(* IEC 61131-3 sources: daoli-st-library/DL_Device (part 32) *)

(* ---- FB_DL_StarDeltaMotor.st ---- *)
(*==============================================================================
 * 组件名称 (Component)  : FB_DL_StarDeltaMotor
 * 所属子库 (Sublibrary) : DL_Device
 * 当前版本 (Version)    : 1.0.1
 * 兼容性   (Platform)   : CODESYS 3.5 / TwinCAT 3 / 汇川 InoProShop / Machine Expert
 *                         仅依赖 Standard.library（TON / R_TRIG），零厂商方言
 * 分类     (Category)   : 设备执行器功能块（Function Block，无接口实现）
 * 功能简述 (Function)   : 星三角降压启动电机控制（三接触器）。星形降压启动
 *                         （起动力矩约三分之一）→ 星角切换死区互锁（星线圈
 *                         分断后方允许角线圈吸合）→ 三角形全压运行；三路
 *                         接触器指令-反馈校验窗（拒动保护）、运行失反馈
 *                         脱扣、热继过载锁存、重启抑制冷却（沿用
 *                         FB_DL_DolMotor 参数范式）；星角输出互斥出口
 *                         断言 + 反馈互锁冲突监视；状态机复用既有
 *                         E_DL_MotorState（禁止重定义），ENUM + CASE + ELSE
 *                         兜底。
 * 开源溯源 (Origin)     : 来源标签 lbp-basic-process / lbp-device
 *                         （RAW_NOTES_R6 S-1 + S-5：星三角降压启动时序、
 *                         星角切换死区时间互锁、三接触器反馈校验等行业
 *                         公知工程惯例，公开教学资料，仅借鉴通用工程语义；
 *                         状态机、死区互锁实现、故障码按本库红线独立设计，
 *                         clean-room 未复制源码）。
 * 红线自检 (Redline)    : R1 零全局变量表/外部变量引用 ✓｜R2 零物理 IO 地址 ✓
 *                         R3 纯 IEC 61131-3 ✓｜R4 防越界/互斥断言 ✓
 *                         R5 全变量中英双语同行注释 ✓｜R6 ENUM+CASE+ELSE ✓
 *                         R7 七个定时器/边缘实例主体最前部无条件刷新 ✓
 * 公约遵循 (Convention) : 0.1/R23 本块为纯事件型状态机（BOOL 指令/反馈 +
 *                         TIME 参数，无积分/滤波类连续量同步语义），免首扫，
 *                         无内部初始化标志。
 *                         0.7 故障码段位 16#0003_xxxx：【故障级】0003_0240
 *                         主接触器拒动 / 0003_0241 星接触器拒动 / 0003_0242
 *                         星接触器分断失败（角拒动码位承接，见偏离③）/
 *                         0003_0243 星角互斥冲突 / 0003_0244 运行失反馈
 *                         脱扣 / 0003_0245 过载锁存 / 0003_0246 星角转换
 *                         失败（角接触器窗内未吸合），全部 R15 锁存仅复位
 *                         可清；【信息级】0003_0208 重启抑制期启动拒绝
 *                         （沿用 FB_DL_DolMotor 既有同义码位，终审裁定统
 *                         一双电机族口径；仅写 uErrorId，不进 bFault，0.2
 *                         公约）。
 * 偏离留档 (Deviation)  : 依 R11 头注释留档，共 3 条：
 *                         ① 信息级码：规格原分配 0003_0102，经与子库
 *                           VERSION.md 故障码表核对，R5 已占用 0102~0104
 *                           （AnalogTransmitter）；且重启抑制拒绝语义在
 *                           FB_DL_DolMotor 已有信息级码位 0003_0208——
 *                           终审裁定同库同语义不设双码，本块改用 0208
 *                           （0105 空置不分配），与规格原意"沿用 DolMotor
 *                           口径"完全一致。
 *                         ② 规格中 0003_0242（角接触器拒动）与 0003_0246
 *                           （星角转换失败）对"死区满后角接触器窗内未吸合"
 *                           同事件重叠；本实现将 0246 用于规格明示的角接触
 *                           器窗内未吸合，0242 承接转换窗口内星接触器反馈
 *                           未按时分断（星粘连/拒分）的互锁异常，两码位
 *                           各自可测。
 *                         ③ 重启抑制冷却计时采用 TON（本库 Standard.library
 *                           既有范式，DolMotor 同口径），无 CPU 钟依赖。
 * 修订历史 (Revision)   :
 *   2026-11-15  v1.0.0  首版入库（R6 轮 · DL_Device 阀门/驱动族深化）
 *   2026-11-15  v1.0.1  终审修复【逻辑级】重启抑制信息级码双码归一：原分配
 *                       0003_0105 与 FB_DL_DolMotor 既有同义码 0003_0208
 *                       重复（同库同语义双码会致 HMI 报警分组重复映射），
 *                       改用 0208 统一口径。引脚契约零变更。
 *============================================================================*)
FUNCTION_BLOCK FB_DL_StarDeltaMotor
VAR_INPUT
    bCmdStart        : BOOL;            // 启动指令（Start command），上升沿生效 / Start command, rising edge effective
    bCmdStop         : BOOL;            // 停止指令（Stop command），电平生效 / Stop command, level effective
    bFbMain          : BOOL;            // 主接触器反馈（Main contactor feedback），TRUE=吸合 / Main contactor feedback, TRUE = picked up
    bFbStar          : BOOL;            // 星形接触器反馈（Star contactor feedback），TRUE=吸合 / Star contactor feedback, TRUE = picked up
    bFbDelta         : BOOL;            // 三角形接触器反馈（Delta contactor feedback），TRUE=吸合 / Delta contactor feedback, TRUE = picked up
    bThermalOverload : BOOL;            // 热继电器过载信号（Thermal overload trip），TRUE=过载 / Thermal overload trip, TRUE = overloaded
    bPermitStart     : BOOL;            // 启动允许联锁（Start permit），TRUE=允许 / Start permit interlock, TRUE = start allowed
    tStarTime        : TIME := T#5S;    // 星形运行时间（Star run time），按负载实测加速时间整定 / Star run time, tune per measured load acceleration
    tDeadTime        : TIME := T#100MS; // 星角转换死区时间（Transition dead time），域 50~200MS，星分断后角方可吸合 / Transition dead time 50..200 ms, star must drop before delta picks up
    tFbWindow        : TIME := T#500MS; // 指令-反馈校验窗口（Feedback check window），T#0S=免校验 / Feedback check window, T#0S disables the check
    tRestartInhibit  : TIME := T#60S;   // 重启抑制冷却时间（Restart inhibit），停机后冷却期内拒绝启动 / Restart inhibit cooling time after stop
    bReset           : BOOL;            // 故障复位（Fault reset），上升沿生效 / Fault reset, rising edge effective
END_VAR

VAR_OUTPUT
    bMainContactor   : BOOL;            // 主接触器线圈输出（Main contactor coil），星形与运行期全程吸合 / Main contactor coil, closed through star and run phases
    bStarContactor   : BOOL;            // 星形接触器线圈输出（Star contactor coil），仅星形降压段吸合 / Star contactor coil, closed only in star phase
    bDeltaContactor  : BOOL;            // 三角形接触器线圈输出（Delta contactor coil），死区满后吸合 / Delta contactor coil, closed after dead time
    eState           : E_DL_MotorState; // 当前状态机状态（Current state），复用既有枚举 / Current state, reuses existing enum
    bRunning         : BOOL;            // 运行反馈（Running feedback），角接触器吸合确认 / Running feedback, confirmed by delta contactor
    bFault           : BOOL;            // 故障锁存中（Fault latched），TRUE=需复位（含过载脱扣）/ Fault latched, TRUE requires reset (incl. overload trip)
    uErrorId         : UDINT;           // 末次故障码（Last error code），0=无故障，段位 16#0003_xxxx / Last error code, 0 = none, family 16#0003_xxxx
    bRestartInhibit  : BOOL;            // 重启抑制激活中（Restart inhibit active），TRUE=冷却期拒绝启动 / Restart inhibit active, TRUE = starts refused
    bStarPhase       : BOOL;            // 星形阶段指示（Star phase active），调试/HMI 用 / Star phase indicator for debug and HMI
    uStartCount      : UDINT;           // 累计启动次数（Start count），每次受理启动 +1 / Total start count, incremented per accepted start
END_VAR

VAR
    _eState           : E_DL_MotorState := E_DL_MotorState.eIdle; // 内部状态机步序（Internal state step）/ Internal state step
    _bFaultLatch      : BOOL;           // 故障锁存标志（Fault latch flag），仅复位清除 / Fault latch flag, cleared only by reset
    _uErrorIdInt      : UDINT;          // 内部故障码寄存（Internal error register），故障级与信息级共用 / Internal error register, fault and info codes share it
    _bDeadZone        : BOOL;           // 星角转换死区子相位（Star-delta dead-zone sub-phase），星形态内二段 / Dead-zone sub-phase inside starting state
    _bDeltaCmd        : BOOL;           // 角接触器指令已发出（Delta command issued），转换校验窗运行中 / Delta command issued, check window running
    _bCooling         : BOOL;           // 冷却计时进行中（Cooling timing active）/ Cooling timer run request flag
    _bRestartInhAct   : BOOL;           // 重启抑制激活内部寄存（Internal restart inhibit register）/ Internal restart inhibit register
    _bFbWinEn         : BOOL;           // 反馈校验窗使能（Feedback window enable），窗口参数大于零有效 / Feedback window enable, active when window above zero
    _bInFbWin         : BOOL;           // 主/星反馈窗计时条件（Main/star window timing condition）/ Timing condition of main and star window
    _bInStarTime      : BOOL;           // 星形运行计时条件（Star run timing condition）/ Timing condition of star run timer
    _bInDeadTime      : BOOL;           // 死区计时条件（Dead time timing condition）/ Timing condition of dead time timer
    _bInDeltaWin      : BOOL;           // 角反馈窗计时条件（Delta window timing condition）/ Timing condition of delta window
    _bInRunningSt     : BOOL;           // 运行态判定中间量（Running-state test intermediate） / Running-state test intermediate
    _fbTrigStart      : R_TRIG;         // 引脚启动指令上升沿（Pin start command edge）/ Pin start command rising edge
    _fbTrigReset      : R_TRIG;         // 引脚复位上升沿（Pin reset edge）/ Pin reset rising edge
    _fbTonFbWin       : TON;            // 主/星接触器反馈校验窗定时器（Main and star feedback window timer）/ Main and star feedback window timer
    _fbTonStarTime    : TON;            // 星形运行时间定时器（Star run time timer）/ Star run time timer
    _fbTonDeadTime    : TON;            // 星角转换死区定时器（Transition dead time timer）/ Transition dead time timer
    _fbTonDeltaWin    : TON;            // 角接触器反馈校验窗定时器（Delta feedback window timer）/ Delta feedback window timer
    _fbTonRestartInh  : TON;            // 重启抑制冷却定时器（Restart inhibit cooling timer）/ Restart inhibit cooling timer
END_VAR

// ============================================================================
// 段 1｜定时器与边缘检测实例无条件周期刷新（R7：严禁置于 IF/CASE 分支内）
//      Unconditional per-cycle refresh of all timer and edge instances (R7)
// ============================================================================
_fbTrigStart(CLK := bCmdStart);
_fbTrigReset(CLK := bReset);
_bFbWinEn := (tFbWindow > T#0S);      // 窗口为零 = 免校验（Zero window = check disabled）
_bInFbWin := (_eState = E_DL_MotorState.eStarting) AND (NOT _bDeadZone) AND _bFbWinEn; // 启动段主/星校验窗（Starting phase main and star window）
_bInStarTime := (_eState = E_DL_MotorState.eStarting) AND (NOT _bDeadZone); // 星形段计时（Star phase timing）
_bInDeadTime := (_eState = E_DL_MotorState.eStarting) AND _bDeadZone AND (NOT _bDeltaCmd); // 死区段计时（Dead-zone timing）
_bInDeltaWin := (_eState = E_DL_MotorState.eStarting) AND _bDeadZone AND _bDeltaCmd AND (NOT bFbDelta) AND _bFbWinEn; // 角校验窗（Delta check window）
_fbTonFbWin(IN := _bInFbWin, PT := tFbWindow);
_fbTonStarTime(IN := _bInStarTime, PT := tStarTime);
_fbTonDeadTime(IN := _bInDeadTime, PT := tDeadTime);
_fbTonDeltaWin(IN := _bInDeltaWin, PT := tFbWindow);
_fbTonRestartInh(IN := _bCooling, PT := tRestartInhibit);

// 冷却到期：解除抑制（Cooling expired: release inhibit）
IF _fbTonRestartInh.Q THEN
    _bCooling       := FALSE;         // 结束冷却计时（Stop cooling timing）
    _bRestartInhAct := FALSE;         // 解除抑制（Release inhibit）
ELSE
    _bRestartInhAct := _bCooling;     // 冷却期间抑制有效（Inhibit active during cooling）
END_IF
_bInRunningSt := (_eState = E_DL_MotorState.eRunning); // 运行态判定（Running-state test）

// ============================================================================
// 段 2｜星角反馈互锁冲突全局监视（优先级最高）：双反馈同真物理不可能
//      Star-delta feedback conflict monitor (highest priority): both
//      feedbacks ON is physically impossible
// ============================================================================
IF bFbStar AND bFbDelta THEN
    _bFaultLatch := TRUE;             // 反馈冲突锁存（Feedback conflict latch）
    _uErrorIdInt := 16#0003_0243;     // 0003_0243 星角互斥冲突【故障级】/ Star-delta exclusivity conflict, fault level
    _eState      := E_DL_MotorState.eFault; // 强制故障态（Force fault state）
END_IF

// ============================================================================
// 段 3｜过载全局监视：启动/运行态过载立即锁存脱扣
//      Global overload monitor: trip immediately in starting/running states
// ============================================================================
IF bThermalOverload AND ((_eState = E_DL_MotorState.eStarting) OR _bInRunningSt) THEN
    _bFaultLatch := TRUE;             // 过载锁存（Overload latched）
    _uErrorIdInt := 16#0003_0245;     // 0003_0245 热继电器过载脱扣【故障级】/ Thermal overload trip, fault level
    _eState      := E_DL_MotorState.eTripOverload; // 强制脱扣态（Force trip state）
END_IF

// ============================================================================
// 段 4｜核心状态机（ENUM + CASE，含 ELSE 非法状态兜底）
//      Core state machine (ENUM + CASE with ELSE illegal-state fallback)
// ============================================================================
CASE _eState OF

    E_DL_MotorState.eIdle: // 空闲停机态：三线圈全断，评估启动请求
        IF _fbTrigStart.Q THEN
            IF bThermalOverload THEN
                // 过载未复位：静默拒绝（Overload present: silent refusal）
            ELSIF NOT bPermitStart THEN
                // 联锁未满足：静默拒绝（Permit absent: silent refusal）
            ELSIF _bRestartInhAct THEN
                _uErrorIdInt := 16#0003_0208; // 0003_0208 重启抑制期内启动被拒【信息级】（沿用 DolMotor 既有同义码位，终审裁定）/ Start refused during restart inhibit, info level (DolMotor shared code, audit ruling)
            ELSE
                _bDeadZone   := FALSE;   // 复位转换子相位（Reset transition sub-phase）
                _bDeltaCmd   := FALSE;   // 复位角指令标志（Reset delta command flag）
                uStartCount  := uStartCount + 1; // 累计启动 +1（Total starts +1）
                _eState      := E_DL_MotorState.eStarting;
            END_IF
        END_IF

    E_DL_MotorState.eStarting: // 启动校验态：星形降压段 → 死区段 → 角校验段
        IF bCmdStop THEN
            _eState := E_DL_MotorState.eStopping; // 停止指令：三线圈全断（Stop: all coils off）
        ELSIF (NOT _bDeadZone) AND (NOT bFbMain) AND _bFbWinEn AND _fbTonFbWin.Q THEN
            _bFaultLatch := TRUE;                 // 主接触器拒动锁存（Main refusal latch）
            _uErrorIdInt := 16#0003_0240;         // 0003_0240 主接触器拒动（窗内未吸合）【故障级】/ Main contactor refused, fault level
            _eState      := E_DL_MotorState.eFault;
        ELSIF (NOT _bDeadZone) AND (NOT bFbStar) AND _bFbWinEn AND _fbTonFbWin.Q THEN
            _bFaultLatch := TRUE;                 // 星接触器拒动锁存（Star refusal latch）
            _uErrorIdInt := 16#0003_0241;         // 0003_0241 星接触器拒动（窗内未吸合）【故障级】/ Star contactor refused, fault level
            _eState      := E_DL_MotorState.eFault;
        ELSIF (NOT _bDeadZone) AND _fbTonStarTime.Q THEN
            _bDeadZone := TRUE;                   // 星形时间计满，星线圈分断，进入死区（Star time elapsed, star coil drops, dead zone entered）
        ELSIF _bDeadZone AND (NOT _bDeltaCmd) AND _fbTonDeadTime.Q THEN
            IF bFbStar THEN
                _bFaultLatch := TRUE;             // 星接触器分断失败锁存（Star drop-out failure latch）
                _uErrorIdInt := 16#0003_0242;     // 0003_0242 星接触器分断失败（死区满仍吸合）【故障级】/ Star contactor failed to drop, fault level
                _eState      := E_DL_MotorState.eFault;
            ELSE
                _bDeltaCmd := TRUE;               // 死区满且星已分断，发出角指令（Dead time done, star dropped, delta commanded）
            END_IF
        ELSIF _bDeadZone AND _bDeltaCmd AND bFbDelta AND (NOT bFbStar) THEN
            _eState := E_DL_MotorState.eRunning;  // 角吸合确认，转全压运行（Delta picked up, to full-voltage running）
        ELSIF _bDeadZone AND _bDeltaCmd AND (NOT bFbDelta) AND _bFbWinEn AND _fbTonDeltaWin.Q THEN
            _bFaultLatch := TRUE;                 // 星角转换失败锁存（Transition failure latch）
            _uErrorIdInt := 16#0003_0246;         // 0003_0246 星角转换失败（角接触器窗内未吸合）【故障级】/ Star-delta transition failed, fault level
            _eState      := E_DL_MotorState.eFault;
        END_IF

    E_DL_MotorState.eRunning: // 全压运行态：主+角吸合确认
        IF bCmdStop THEN
            _eState := E_DL_MotorState.eStopping; // 停止指令（Stop command）
        ELSIF (NOT bFbDelta) OR (NOT bFbMain) THEN
            _bFaultLatch := TRUE;                 // 失反馈脱扣锁存（Feedback loss latch）
            _uErrorIdInt := 16#0003_0244;         // 0003_0244 运行中反馈意外断开【故障级】/ Contactor feedback dropped while running, fault level
            _eState      := E_DL_MotorState.eFault;
        END_IF

    E_DL_MotorState.eStopping: // 停机过渡态：三线圈已断，等反馈全部分断
        IF (NOT bFbMain) AND (NOT bFbStar) AND (NOT bFbDelta) THEN
            _bDeadZone := FALSE;                  // 复位转换子相位（Reset transition sub-phase）
            _bDeltaCmd := FALSE;                  // 复位角指令标志（Reset delta command flag）
            _bCooling  := TRUE;                   // 启动重启抑制冷却（Start restart-inhibit cooling）
            _eState    := E_DL_MotorState.eIdle;  // 回空闲（Back to idle）
        END_IF
        // 反馈触点粘连时保持本态等待分断，直至上层干预（Welded contacts hold this state until intervention）

    E_DL_MotorState.eTripOverload: // 过载脱扣锁存态：仅复位且过载消失后可清
        IF _fbTrigReset.Q AND (NOT bThermalOverload) THEN
            _bFaultLatch := FALSE;                // 解除锁存（Release latch）
            _uErrorIdInt := 0;                    // 故障码清零（Error code cleared）
            _bDeadZone   := FALSE;                // 复位转换子相位（Reset transition sub-phase）
            _bDeltaCmd   := FALSE;                // 复位角指令标志（Reset delta command flag）
            _bCooling    := TRUE;                 // 脱扣复位后同样进入冷却（Cooling also after trip reset）
            _eState      := E_DL_MotorState.eIdle; // 回空闲（Back to idle）
        END_IF

    E_DL_MotorState.eFault: // 故障锁存态：仅复位可退出
        IF _fbTrigReset.Q THEN
            _bFaultLatch := FALSE;                // 解除锁存（Release latch）
            _uErrorIdInt := 0;                    // 故障码清零（Error code cleared）
            _bDeadZone   := FALSE;                // 复位转换子相位（Reset transition sub-phase）
            _bDeltaCmd   := FALSE;                // 复位角指令标志（Reset delta command flag）
            _bCooling    := TRUE;                 // 故障复位后进入冷却（Cooling also after fault reset）
            _eState      := E_DL_MotorState.eIdle; // 回空闲（Back to idle）
        END_IF

    ELSE // 非法状态兜底：任何越界枚举值强制锁存故障（Illegal state fallback）
        _bFaultLatch := TRUE;                     // 故障锁存（Fault latched）
        _uErrorIdInt := 16#0003_0201;             // 0003_0201 非法状态【故障级】（沿用库级既有码）/ Illegal state, fault level
        _eState      := E_DL_MotorState.eFault;
END_CASE

// ============================================================================
// 段 5｜线圈输出推导 + 星角互斥出口断言（硬约束：星/角输出恒不可同真）
//      Coil output derivation + star-delta exclusivity exit assertion
// ============================================================================
bMainContactor  := (_eState = E_DL_MotorState.eStarting) OR (_eState = E_DL_MotorState.eRunning); // 启动段与运行段主接触器吸合（Main closed in starting and running）
bStarContactor  := (_eState = E_DL_MotorState.eStarting) AND (NOT _bDeadZone); // 仅星形降压段吸合（Closed only in star phase）
bDeltaContactor := (_eState = E_DL_MotorState.eRunning);       // 仅全压运行段吸合（Closed only in full-voltage run）
IF bStarContactor AND bDeltaContactor THEN
    bStarContactor  := FALSE;                        // 断言对调：异常同真时双断保安全（Assertion fallback: cut both on impossible condition）
    bDeltaContactor := FALSE;
    _bFaultLatch    := TRUE;                         // 出口冲突锁存（Exit conflict latch）
    _uErrorIdInt    := 16#0003_0243;                 // 0003_0243 星角互斥冲突【故障级】/ Star-delta exclusivity conflict, fault level
    _eState         := E_DL_MotorState.eFault;
END_IF

// ============================================================================
// 段 6｜状态引脚映射（bFault 为显式派生式，排除信息级码——0.2 公约）
//      Status pin mapping (bFault explicit derived form, info codes excluded)
// ============================================================================
eState          := _eState;                        // 状态映射（State mapping）
bRunning        := (_eState = E_DL_MotorState.eRunning) AND bFbDelta; // 运行 = 状态且角接触器确认（Running = state AND delta confirmed）
bFault          := _bFaultLatch OR (_eState = E_DL_MotorState.eFault) OR (_eState = E_DL_MotorState.eTripOverload); // 故障派生（Fault derived）
uErrorId        := _uErrorIdInt;                   // 故障码映射（Error code mapping）
bRestartInhibit := _bRestartInhAct;                // 重启抑制映射（Restart inhibit mapping）
bStarPhase      := (_eState = E_DL_MotorState.eStarting) AND (NOT _bDeadZone); // 星形阶段指示（Star phase indicator）
END_FUNCTION_BLOCK

(* ---- FB_DL_SteamTrapSurvey.st ---- *)
(*==============================================================================
 * 组件名称 (Component)  : FB_DL_SteamTrapSurvey
 * 所属子库 (Sublibrary) : DL_Device
 * 当前版本 (Version)    : 1.0.0
 * 兼容性 (Platform)     : CODESYS 3.5+ / TwinCAT 3 / 汇川 InoProShop / 施耐德 Machine Expert
 *                         仅依赖 Standard.library（TON / ABS），零厂商私有库
 * 功能描述 (Function)   : 疏水阀温度周期特征普查与失效分级。对单阀（多实例
 *                         部署即跨管网普查）滚动窗（tCycleWin 自复位 TON）内
 *                         累计阀温-环境温差样本，窗到时按平均温差分级：
 *                         >= fDTOpen 判直通泄漏（eLeak）、<= fDTClosed 判
 *                         堵塞冷阀（eBlock）、介于其间健康（eOk）。与
 *                         SteamTrapMonitor/DiagTrend（单阀监测与温差趋势）
 *                         分工：本件是周期窗普查 + 失效分级的语义。
 * 来源标签 (Origin)     : ROADMAP §21.5 R13 池（L920），自研 clean-room
 * 边界语义 (Boundary)   : ① 温度 NaN/Inf 拍拒收（不入累计不推进计数）；
 *                         ② 滚动窗 TON 自复位（IN 带 NOT tonWin.Q，FB33-2），
 *                         窗到时单拍清累计（真滚动窗口径）；
 *                         ③ 分级门限配比约束 fDTOpen > fDTClosed（组态闸）；
 *                         ④ 窗未满最小样本数（nMinSamp）不判级（防短窗误报）。
 * 输出语义 (Fallback)   : 【R191】bEnable = FALSE → 分级保持末值 + 测量出口
 *                         FALSE（普查监视失能必须收敛）；eFault 相 → 冻结
 *                         + bError = TRUE。
 * 码位     (Codes)      : 按 R297 范式零 16# 码位硬编码；错误出口 BOOL+ENUM(eCause)。
 * 红线自检 (Redline)    : 7 项红线已自检：R1 零全局 ✓｜R2 零物理地址 ✓｜R3 纯 IEC ✓
 *                         R4 除零（计数 eps 闸）/NaN 拒收/组态闸 ✓｜R5 双语同行注释 ✓
 *                         R6 CASE 带 ELSE 兜底迁 eFault ✓｜R7 TON/R_TRIG 段 0 无条件刷新 ✓
 * 验收向量 (Acceptance) : V1 窗内温差均值 45（fDTOpen=30）→ eHealth=eLeak；
 *                         V2 均值 5（fDTClosed=10）→ eHealth=eBlock；
 *                         V3 均值 20 → eHealth=eOk；V4 窗内样本 < 8 →
 *                         eHealth=eUnknown 不判级。
 * 修订历史 (Revision)   : 2026-11-20  v1.0.0  R51 首版（批 3 · 序号 14）
 *==============================================================================*)
TYPE E_DL_StsHealth :
(
    eOk      := 0,                           (* 健康（温差居中带） / Healthy *)
    eLeak    := 1,                           (* 直通泄漏（温差持续高） / Steam leaking *)
    eBlock   := 2,                           (* 堵塞冷阀（温差持续低） / Blocked cold trap *)
    eUnknown := 3                            (* 样本不足未判级 / Insufficient samples *)
);
END_TYPE

TYPE E_DL_StsState :
(
    eIdle  := 0,                             (* 待使能 / Idle *)
    eSurvey:= 10,                            (* 普查运行 / Survey run *)
    eFault := 90                             (* 故障锁存相 / Fault latched phase *)
);
END_TYPE

TYPE E_DL_StsCause :
(
    eNone       := 0,                        (* 无故障成因 / No cause *)
    eCfgIllegal := 1,                        (* 组态非法：窗时/门限/秒值越域 / Illegal config *)
    ePhaseBad   := 2                         (* 非法相位兜底 / Illegal phase fallback *)
);
END_TYPE

FUNCTION_BLOCK FB_DL_SteamTrapSurvey
VAR_INPUT
    fTempC     : LREAL := 0.0;               (* 阀体温度 [°C] / Trap body temperature *)
    fAmbC      : LREAL := 25.0;              (* 环境参考温度 [°C] / Ambient reference *)
    tCycleWin  : TIME := T#60S;              (* 普查滚动窗时长，域 > T#0S [ms] / Survey window time *)
    fDTOpen    : LREAL := 30.0;              (* 直通泄漏门限（均值 >= 判泄），域 > fDTClosed [K] / Leak threshold *)
    fDTClosed  : LREAL := 10.0;              (* 堵塞冷阀门限（均值 <= 判堵），域 < fDTOpen [K] / Block threshold *)
    nMinSamp   : INT := 8;                   (* 判级最小样本数，域 1..999 [点] / Min samples for verdict *)
    fScanS     : LREAL := 1.0;               (* 扫描周期秒值，域 > 1E-6 [s] / Scan period seconds *)
    bEnable    : BOOL := TRUE;               (* 使能 [-] / Enable *)
    bReset     : BOOL := FALSE;              (* 复位命令，上升沿清全部 [-] / Reset command *)
END_VAR
VAR_OUTPUT
    fDtAvg     : LREAL;                      (* 最近窗平均温差 [K] / Window mean delta-T *)
    eHealth    : E_DL_StsHealth;             (* 失效分级出口（信息级逐窗重算，R189） / Health grade outlet *)
    nSampCnt   : INT;                        (* 最近窗样本数 [点] / Window sample count *)
    bWinTick   : BOOL;                       (* 窗到时单拍脉冲 [-] / Window expiry pulse *)
    eState     : E_DL_StsState;              (* 状态出口 / State outlet *)
    eCause     : E_DL_StsCause;              (* 故障成因出口 / Fault cause outlet *)
    bError     : BOOL;                       (* 故障锁存标志 [-] / Fault latch flag *)
END_VAR
VAR
    _eState  : E_DL_StsState := E_DL_StsState.eIdle;      (* 内部相位（CASE 唯一写入目标） / Internal phase *)
    _eCause  : E_DL_StsCause := E_DL_StsCause.eNone;      (* 故障成因锁存量 / Latched cause *)
    rtReset  : R_TRIG;                       (* 复位沿实例，段 0 无条件调用 / Reset edge instance *)
    tonWin   : TON;                          (* 普查滚动窗自复位计时，段 0 无条件调用 / Self-resetting survey window *)
    _fDtSum  : LREAL;                        (* 窗内温差累计 [K] / Delta-T window sum *)
    _fDt     : LREAL;                        (* 本拍温差派生量 [K] / Delta-T this scan *)
    _nSamp   : INT;                          (* 窗样本计数 [点] / Window sample count *)
    _nSampMax: INT;                          (* 窗样本计数上限锁存（防 INT 溢出）[点] / Sample cap latch *)
    _fAvg    : LREAL;                        (* 窗均值工作量 [K] / Window mean work *)
    _bTick   : BOOL;                         (* 窗到时单拍量 [-] / Window tick work *)
    _bTempBad: BOOL;                        (* 温度非有限当拍量 [-] / Non-finite temperature *)
    _bFault  : BOOL;                         (* 故障锁存位 / Latched fault bit *)
    _bCfgBad : BOOL;                         (* 组态非法当拍量 / Illegal config this scan *)
END_VAR
VAR CONSTANT
    DL_STS_EPS  : LREAL := 1.0E-6;           (* 秒值/计数判零容差 [-] / Epsilon *)
    DL_STS_NCAP : INT   := 999;              (* 窗样本计数上限（防 INT 溢出）[点] / Sample cap *)
END_VAR

(* —— 段 0：当拍判据派生 + 实例无条件刷新（R228A） —— *)
_bCfgBad := (tCycleWin <= T#0S) OR (fDTOpen <= fDTClosed) OR (nMinSamp < 1) OR (nMinSamp > DL_STS_NCAP)
            OR (fScanS <= DL_STS_EPS);   (* 组态闸（R151 全引脚 + 门限序 R146） / Config gate *)
rtReset(CLK := bReset);                      (* 复位沿每拍必调 / Reset edge every scan *)
_bTempBad := (fTempC <> fTempC) OR ((fTempC - fTempC) <> (fTempC - fTempC))
            OR (fAmbC <> fAmbC) OR ((fAmbC - fAmbC) <> (fAmbC - fAmbC));   (* 双温度 NaN 自反 + Inf 差判 / Non-finite temperature gates *)
tonWin(IN := (_eState = E_DL_StsState.eSurvey) AND NOT tonWin.Q, PT := tCycleWin);   (* 滚动窗自复位计时（FB33-2） / Self-resetting window *)
_bTick := tonWin.Q;                          (* 窗到时单拍量 / Window tick work *)

(* —— 段 1：单拍量预清零（R107） —— *)
_fDt := 0.0;                                 (* 温差预清（每拍全路径派生，R285） / Delta-T preset *)
_fAvg := 0.0;                                (* 均值预清 / Mean preset *)
bWinTick := FALSE;                           (* 窗到时脉冲预清，唯一分支置位 / Tick preset *)
_nSampMax := DL_STS_NCAP;                    (* 计数上限预置 / Cap preset *)

(* —— 段 2：复位沿处理（作用域：清故障 + 清窗累计 + 清样本计数 + 清分级出口 + 迁 eIdle，R283 逐项声明） —— *)
IF rtReset.Q THEN
    _bFault := FALSE;                        (* 清故障锁存 / Clear fault *)
    _eCause := E_DL_StsCause.eNone;          (* 清成因 / Clear cause *)
    _fDtSum := 0.0;                          (* 清窗累计 / Clear sum *)
    _nSamp := 0;                             (* 清样本计数 / Clear count *)
    fDtAvg := 0.0;                           (* 清均值出口 / Clear mean outlet *)
    eHealth := E_DL_StsHealth.eUnknown;      (* 分级回未知 / Grade unknown *)
    nSampCnt := 0;                           (* 清样本出口 / Clear count outlet *)
    _eState := E_DL_StsState.eIdle;          (* 迁待机相 / Back to idle *)
END_IF

(* —— 段 3：组态闸故障锁存（R45 配对；锁存至复位沿，R189） —— *)
IF _bCfgBad AND NOT _bFault THEN
    _bFault := TRUE;                         (* 锁存故障位 / Latch fault *)
    _eCause := E_DL_StsCause.eCfgIllegal;    (* 成因：组态非法 / Cause: illegal config *)
    _eState := E_DL_StsState.eFault;         (* 同步迁故障相 / Migrate to fault *)
END_IF

(* —— 段 4：CASE 主状态机（ELSE 兜底迁 eFault，红线 6） —— *)
CASE _eState OF
    E_DL_StsState.eIdle:                     (* 待机相 / Idle *)
        IF bEnable AND NOT _bFault AND NOT _bTempBad THEN
            _eState := E_DL_StsState.eSurvey;   (* 进入普查 / Enter survey *)
        END_IF
    E_DL_StsState.eSurvey:                   (* 普查相：滚动窗累计 + 到时分级 / Survey *)
        IF NOT bEnable THEN
            _eState := E_DL_StsState.eIdle;  (* 失能回待机（分级保持末值，R191 声明） / Back to idle *)
        ELSE
            IF NOT _bTempBad THEN
                _fDt := fTempC - fAmbC;      (* 温差派生（减法无除零） / Delta-T derive *)
                _fDtSum := _fDtSum + _fDt;   (* 窗累计 / Sum into window *)
                IF _nSamp < _nSampMax THEN
                    _nSamp := _nSamp + 1;    (* 样本计数（上限内防 INT 溢出） / Count sample *)
                END_IF
            END_IF                           (* 温度坏值拍：拒收不入累计（边界①） / Bad scan: reject *)
            IF _bTick THEN                   (* 窗到时单拍：分级 + 清窗（滚动窗口径，边界②） / On window tick *)
                bWinTick := TRUE;            (* 窗到时脉冲 / Tick pulse *)
                nSampCnt := _nSamp;          (* 窗样本数出口快照 / Count snapshot *)
                IF _nSamp >= nMinSamp THEN   (* 最小样本闸（边界④） / Min-sample gate *)
                    _fAvg := _fDtSum / INT_TO_LREAL(_nSamp);   (* 窗均值（除子 >= nMinSamp >= 1，无除零） / Window mean *)
                    fDtAvg := _fAvg;         (* 均值出口刷新 / Mean outlet *)
                    IF _fAvg >= fDTOpen THEN
                        eHealth := E_DL_StsHealth.eLeak;   (* 直通泄漏（独立分级，R190） / Leak grade *)
                    ELSIF _fAvg <= fDTClosed THEN
                        eHealth := E_DL_StsHealth.eBlock;  (* 堵塞冷阀（独立分级） / Block grade *)
                    ELSE
                        eHealth := E_DL_StsHealth.eOk;     (* 健康居中带（IF 链 ELSE 兜底，R285） / Healthy *)
                    END_IF
                ELSE
                    eHealth := E_DL_StsHealth.eUnknown;   (* 样本不足未判级 / Unknown *)
                    fDtAvg := 0.0;           (* 未判级均值出口回哨兵 / Mean sentinel *)
                END_IF
                _fDtSum := 0.0;              (* 清窗累计（下一窗起算） / Clear sum *)
                _nSamp := 0;                 (* 清样本计数 / Clear count *)
            END_IF
        END_IF
    E_DL_StsState.eFault:                    (* 故障相：冻结保持，仅复位沿出 / Fault *)
        ;                                    (* 锁存回放（R28） / Replay from latch *)
    ELSE                                     (* 非法相位兜底迁安全态 / Illegal phase fallback *)
        _eState := E_DL_StsState.eFault;     (* 迁故障相 / To fault *)
        _bFault := TRUE;                     (* 同步锁存 / Latch *)
        _eCause := E_DL_StsCause.ePhaseBad;  (* 成因：非法相位 / Cause: illegal phase *)
END_CASE

(* —— 段 5：出口映射（bError/eState 同源，R191） —— *)
bWinTick := _bTick;                          (* 窗到时脉冲出口 / Tick outlet *)
bError := _bFault;                           (* 故障标志镜像 / Fault flag mirror *)
eState := _eState;                           (* 状态出口 / State outlet *)
eCause := _eCause;                           (* 成因出口 / Cause outlet *)
END_FUNCTION_BLOCK

(* ---- FB_DL_StepperMicroFeedPulseEquiv.st ---- *)
//==============================================================================
// 功能块：FB_DL_StepperMicroFeedPulseEquiv ｜ 中文名称：步进细分脉冲当量换算与组态校验
// 所属子库：DL_Device ｜ 版本：v1.0.0 ｜ 兼容：CODESYS V3.5+ / TwinCAT 3 / 汇川 InoProShop
// 功能描述：步进电机细分脉冲当量链换算——整步数 x 细分数 x 减速比 / 丝距
//           导程 → 脉冲当量（脉冲/mm 与 mm/脉冲），并按反向间隙换算补偿
//           脉冲数；组态域校验复用 FB_DL_PulseDirStepper 的组态纪律
//           （细分 1..256 整数、导程/整步数/减速比 > 0）。触发式：bExecute
//           上升沿启动计算，结果锁存至下次触发或复位。细分数非 2 的幂
//           按实际值照算并给信息级提示（驱动器只认 2 的幂档位时由
//           上层拦截，本件不阻断换算链可观测性）。
// 开源溯源 (Origin)：道莅原创实现（参考步进驱动细分与丝距传动工程惯例 分类与参数域）
// 单位表：整步数[步/转] / 细分数[倍] / 减速比[倍] / 导程[毫米每转] /
//         脉冲当量[脉冲每毫米] / 间隙[毫米] / 时间[ms]
// 错误码表：16#0003_0186 信息级（细分数非 2 的幂，按实际值照算，不置
//           bError）/ 16#0003_0187 信息级（反向间隙组态为 0，无间隙补偿
//           提请确认，不置 bError）/ 16#0003_035A 故障级（导程/整步数/
//           减速比 <= 0 或任一输入非有限，组态非法，置 bError）/
//           16#0003_035B 故障级（细分数 <= 0、> 256 或非整数，组态域
//           校验失败，置 bError——该场景不可由 035A 的比值类判据观测，
//           属细分数独立域） / 16#0003_035C 故障级兜底（状态机落 ELSE
//           或非法状态，置 bError）
// 状态机：E_DL_StepperEquivState（四态：eIdle=0 / eCalc=10 / eDone=20 /
//           eFault=99），CASE 含 ELSE 兜底，ELSE 置 035C 并冻结输出
// 边界行为：① 组态非法（035A/035B）→ 进故障态，输出冻结为零，bReset
//           复位；② 细分数非 2 的幂但域内整数 → 照算 + 信息 0186；
//           ③ 间隙为 0 → 照算 + 信息 0187（合法但提请确认）；
//           ④ eDone 态结果锁存保持，新触发沿才重算（防每拍抖动）；
//           ⑤ 失能（bExecute 撤销）不回零——当量是组态量非过程量，
//           锁存保持直至复位；⑥ 安全侧 = 故障态输出全零，禁止残当量
//           进入下游脉冲换算。
// 依赖纪律：Device 域组态件，复用 FB_DL_PulseDirStepper 组态纪律（域值
//           一致性由本件头注释承担验证责任，改动任一侧须复核另一侧）。
// 修订历史：v1.0.0 2026-11-17 首版（R24 派单 · ROADMAP P2 §588）
//==============================================================================

(*------------------------------------------------------------------------------
 * 枚举: E_DL_StepperEquivState（归属本功能块，同文件发布，全库唯一定义）
 * 含义: 当量计算触发式相位，每个成员在 CASE 中有且仅有一个标签。
 *-----------------------------------------------------------------------------*)
TYPE E_DL_StepperEquivState :
(
    eIdle  := 0,   // 空闲：等触发沿 / Idle, awaiting trigger edge
    eCalc  := 10,  // 计算中：本拍完成换算并转出 / Calculating, conversion completed within this scan
    eDone  := 20,  // 完成：结果锁存保持 / Done, results latched
    eFault := 99   // 故障：组态非法/非法状态 / Fault, illegal config or illegal state
);
END_TYPE

FUNCTION_BLOCK FB_DL_StepperMicroFeedPulseEquiv
VAR_INPUT
    bExecute     : BOOL;                    // 触发计算 [—]，上升沿生效 / Trigger calculation, rising edge
    bReset       : BOOL;                    // 故障复位 [—]，上升沿清故障态 / Fault reset, rising edge clears the fault state
    fStepsPerRev : LREAL := 200.0;          // 整步数 [步每转]，典型 200（1.8 度步距角） / Full steps per revolution [steps/rev], typical 200
    fMicroStep   : LREAL := 16.0;           // 细分数 [倍]，有效域 1..256 整数，非 2 的幂给信息级提示 / Microstepping divisor [count], valid range 1..256 integer
    fGearRatioIn : LREAL := 1.0;            // 减速比（电机转/丝杠转）[倍]，须 > 0 / Gear reduction ratio [ratio], must be > 0
    fLeadMm      : LREAL := 5.0;            // 丝杠导程 [毫米每转]，须 > 0 / Screw lead [mm/rev], must be > 0
    fBacklashMm  : LREAL := 0.0;            // 反向间隙 [毫米]，>= 0，为 0 给信息级提示 / Backlash [mm], >= 0, zero raises an info notice
END_VAR
VAR_OUTPUT
    fPulsePerMm    : LREAL;                 // 脉冲当量 [脉冲每毫米] / Pulse equivalent [pulses/mm]
    fMmPerPulse    : LREAL;                 // 反向当量 [毫米每脉冲] / Inverse equivalent [mm/pulse]
    fBacklashPulse : LREAL;                 // 间隙补偿脉冲数 [脉冲] / Backlash compensation pulses [pulses]
    eState         : E_DL_StepperEquivState; // 相位出口 [—] / Phase outlet
    eErr           : UDINT;                 // 错误码，0 = 无错，码位 16#0003_0186 起信息级、16#0003_035A 起故障级（分带见错误码表） / Error code, 0 = no error, band info/fault per the code table
    bError         : BOOL;                  // 故障级标志，仅故障级错误置位 / Fault-class flag, set only on fault-level codes
    bValid         : BOOL;                  // 输出可用标志 / Outputs usable flag
END_VAR
VAR
    fbTrig       : R_TRIG;                  // 触发沿检测（待机/故障分支同样无条件刷新） / Trigger edge detector, refreshed unconditionally
    _eState      : E_DL_StepperEquivState := E_DL_StepperEquivState.eIdle; // 当前相位 / Current phase
    _bCfgBadA    : BOOL;                    // 035A 类组态非法锁存 / Config fault latch of class 035A
    _bCfgBadB    : BOOL;                    // 035B 类细分数域非法锁存 / Microstep domain fault latch
    _bInfoPow2   : BOOL;                    // 非 2 的幂信息当拍标志 / Non-power-of-two info flag of this scan
    _bInfoNoBl   : BOOL;                    // 间隙为零信息当拍标志 / Zero-backlash info flag of this scan
    _bIllegal    : BOOL;                    // 非法状态标志 / Illegal state flag
    _nMicroDi    : DINT;                    // 细分数整数副本 [倍] / Integer copy of the microstep divisor
    _bInit       : BOOL := FALSE;           // 首扫标志，初值 FALSE 取非判定 / First-scan flag, tested negated
END_VAR
VAR CONSTANT
    DL_SPE_INF      : LREAL := 1.7976931348623157E308; // LREAL 幅值上限 / LREAL magnitude ceiling
    DL_SPE_EPS      : LREAL := 1.0E-6;      // 浮点判零/整判容差 [倍] / Float zero and integrality tolerance [count]
    DL_SPE_MICRO_MAX: LREAL := 256.0;       // 细分数上限 [倍] / Microstep divisor ceiling [count]
    DL_SPE_ZERO     : LREAL := 0.0;         // 零值常量，避免裸字面量 [—] / Zero constant, avoids a bare literal
END_VAR

(*------------------------------------------------------------------------------
 * 段 1｜每拍预置：输出安全侧清零，单拍标志预清零
 *      Outputs cleared fail-safe first, one-shot flags pre-cleared
 *-----------------------------------------------------------------------------*)
fPulsePerMm    := DL_SPE_ZERO;             // 脉冲当量先清（安全侧） / Pulse equivalent cleared first
fMmPerPulse    := DL_SPE_ZERO;             // 反向当量先清 / Inverse equivalent cleared first
fBacklashPulse := DL_SPE_ZERO;             // 间隙脉冲先清 / Backlash pulses cleared first
eErr   := 16#0000_0000;                     // 错误码每拍重算 / Error code recomputed
bError := FALSE;                            // 故障标志每拍重算 / Fault flag recomputed
bValid := FALSE;                            // 可用标志每拍重算 / Usable flag recomputed
_bInfoPow2 := FALSE;                        // 非 2 幂信息预清零 / Power-of-two info pre-cleared
_bInfoNoBl := FALSE;                        // 间隙零信息预清零 / Zero-backlash info pre-cleared
_bIllegal  := FALSE;                        // 非法状态预清零 / Illegal flag pre-cleared

(*------------------------------------------------------------------------------
 * 段 2｜首扫初始化
 *      First-scan initialisation
 *-----------------------------------------------------------------------------*)
IF NOT _bInit THEN
    _eState   := E_DL_StepperEquivState.eIdle; // 相位空闲起步 / Phase starts idle
    _bCfgBadA := FALSE;                     // 组态锁存清零 / Config latch cleared
    _bCfgBadB := FALSE;                     // 细分数锁存清零 / Microstep latch cleared
    _bInit    := TRUE;                      // 首扫只做一次 / The first scan runs once
END_IF

(*------------------------------------------------------------------------------
 * 段 3｜触发沿无条件刷新（R40：CASE 之外每拍必调）
 *      Trigger edge refreshed unconditionally per R40
 *-----------------------------------------------------------------------------*)
fbTrig(CLK := bExecute);                    // 触发沿检测 / Trigger edge detection

(*------------------------------------------------------------------------------
 * 段 4｜组态域校验闸：比值类（035A）与细分数域（035B）分域锁存
 *      Configuration gates in two domains, latched separately
 *-----------------------------------------------------------------------------*)
IF (fLeadMm <> fLeadMm) OR (ABS(fLeadMm) > DL_SPE_INF)
   OR (fStepsPerRev <> fStepsPerRev) OR (ABS(fStepsPerRev) > DL_SPE_INF)
   OR (fGearRatioIn <> fGearRatioIn) OR (ABS(fGearRatioIn) > DL_SPE_INF)
   OR (fBacklashMm <> fBacklashMm) OR (ABS(fBacklashMm) > DL_SPE_INF)
   OR (fMicroStep <> fMicroStep) OR (ABS(fMicroStep) > DL_SPE_INF) THEN
    _bCfgBadA := TRUE;                      // 非有限归入比值类非法（035A） / Non-finite folded into class 035A
END_IF
IF (NOT _bCfgBadA) AND ((fLeadMm <= DL_SPE_EPS) OR (fStepsPerRev <= DL_SPE_EPS)
   OR (fGearRatioIn < DL_SPE_EPS)) THEN
    _bCfgBadA := TRUE;                      // 比值类组态非法锁存（导程/整步数/减速比任一 <= 容差） / Ratio-class config latched
END_IF
IF (NOT _bCfgBadA) AND ((fMicroStep < (DL_SPE_ZERO + DL_SPE_EPS))
   OR (fMicroStep > DL_SPE_MICRO_MAX)) THEN
    _bCfgBadB := TRUE;                      // 细分数域外锁存（035B） / Microstep domain latched
END_IF
IF (NOT _bCfgBadA) AND (NOT _bCfgBadB) THEN
    IF ABS(fMicroStep - LREAL_TO_DINT(fMicroStep)) > DL_SPE_EPS THEN
        _bCfgBadB := TRUE;                  // 细分数非整数锁存（035B） / Non-integer microstep latched
    ELSE
        _nMicroDi := LREAL_TO_DINT(fMicroStep); // 整数副本（域内已闸，转换安全） / Integer copy, range-gated
        IF (_nMicroDi > 1) AND ((_nMicroDi AND (_nMicroDi - 1)) <> 0) THEN
            _bInfoPow2 := TRUE;             // 非 2 的幂：照算并提示（信息级） / Non-power-of-two, computed with an info notice
        END_IF
    END_IF
END_IF
IF (NOT _bCfgBadA) AND (ABS(fBacklashMm) <= DL_SPE_EPS) THEN
    _bInfoNoBl := TRUE;                     // 间隙为 0 提示（信息级） / Zero-backlash notice, info
END_IF

(*------------------------------------------------------------------------------
 * 段 5｜相位机（CASE 含 ELSE 兜底；状态改写只出现在分支判据内，R39）
 *      Phase machine with ELSE fallback, state writes only inside branches
 *-----------------------------------------------------------------------------*)
CASE _eState OF

    E_DL_StepperEquivState.eIdle:          // 空闲：触发沿且组态合法进计算
        IF fbTrig.Q AND (NOT _bCfgBadA) AND (NOT _bCfgBadB) THEN
            _eState := E_DL_StepperEquivState.eCalc; // 进计算相 / To the calc phase
        ELSIF fbTrig.Q AND (_bCfgBadA OR _bCfgBadB) THEN
            _eState := E_DL_StepperEquivState.eFault; // 组态非法进故障 / Illegal config to fault
        END_IF

    E_DL_StepperEquivState.eCalc:          // 计算：本拍完成换算并转完成
        // 拍 N 进入（触发沿且组态合法）/ 本拍行为：换算并锁存 / 拍 N+1 转出：进 eDone 保持
        fPulsePerMm := fStepsPerRev * fMicroStep * fGearRatioIn / fLeadMm; // 脉冲当量 [脉冲每毫米]，分母已闸 / Pulse equivalent, denominator gated
        fMmPerPulse := 1.0 / fPulsePerMm;   // 反向当量 [毫米每脉冲]，分子恒 1 无除零路径 / Inverse equivalent, numerator is 1
        fBacklashPulse := fBacklashMm * fPulsePerMm; // 间隙补偿脉冲 [脉冲] / Backlash compensation pulses
        _eState := E_DL_StepperEquivState.eDone; // 进完成态锁存 / To done, results latched

    E_DL_StepperEquivState.eDone:          // 完成：结果锁存保持，新沿才重算
        IF fbTrig.Q AND (_bCfgBadA OR _bCfgBadB) THEN
            _eState := E_DL_StepperEquivState.eFault; // 组态漂移非法进故障 / Config drift to fault
        ELSIF fbTrig.Q THEN
            _eState := E_DL_StepperEquivState.eCalc; // 新触发沿重算 / New edge recomputes
        END_IF

    E_DL_StepperEquivState.eFault:         // 故障：复位沿且组态恢复合法回空闲
        IF bReset AND (NOT _bCfgBadA) AND (NOT _bCfgBadB) THEN
            _bCfgBadA := FALSE;             // 复位清锁存 / Reset clears the latch
            _bCfgBadB := FALSE;             // 复位清锁存 / Reset clears the latch
            _eState := E_DL_StepperEquivState.eIdle; // 回空闲 / Back to idle
        END_IF

    ELSE                                   // 非法状态兜底（R21：CASE 必带 ELSE）
        _bIllegal := TRUE;                 // 标记非法状态 / Flag the illegal state
        _eState   := E_DL_StepperEquivState.eFault; // 回故障态（输出全零） / Back to fault, outputs zeroed
END_CASE

(*------------------------------------------------------------------------------
 * 段 6｜码位出口与放行（故障级码 3 行内置 bError，R45/R101 配对）
 *      Code outlet and release, fault codes paired with bError
 *-----------------------------------------------------------------------------*)
IF _bIllegal THEN
    eErr   := 16#0003_035C;                 // 故障级：状态机兜底 / Fault: state machine fallback
    bError := TRUE;                         // 置故障标志 / Raise the fault flag
ELSIF _bCfgBadA THEN
    eErr   := 16#0003_035A;                 // 故障级：比值类组态非法 / Fault: ratio-class config illegal
    bError := TRUE;                         // 置故障标志 / Raise the fault flag
ELSIF _bCfgBadB THEN
    eErr   := 16#0003_035B;                 // 故障级：细分数域校验失败 / Fault: microstep domain check failed
    bError := TRUE;                         // 置故障标志 / Raise the fault flag
ELSIF _bInfoPow2 THEN
    eErr := 16#0003_0186;                   // 信息级：细分数非 2 的幂照算 / Info: non-power-of-two divisor, computed as-is
ELSIF _bInfoNoBl THEN
    eErr := 16#0003_0187;                   // 信息级：间隙为 0 提请确认 / Info: zero backlash notice
END_IF

bValid := (NOT bError) AND (_eState = E_DL_StepperEquivState.eDone); // 仅完成态放行 / Usable only in the done phase
eState := _eState;                          // 相位出口 / Phase outlet
END_FUNCTION_BLOCK

(* ---- FB_DL_StrainFatigueCounter.st ---- *)
(* ===========================================================================
   组件名   : FB_DL_StrainFatigueCounter
   分类     : DL_Device / 应变疲劳循环计数
   一句话   : 简化雨流（峰值谷值三点配对）统计循环幅值并累积线性 S-N 损伤度
   复杂度   : 3        版本 : v1.0.0        日期 : 2026-11-24
   开源溯源 : 无（clean-room 自研，未借鉴任何开源实现）
   输入契约 : fStrain 应变输入 [µε]；fDeadBand 反转识别死区 [µε]
              fSnCoeff S-N 系数，即 N=1 对应的循环幅值 [µε]
              fDamageLimit 损伤度限值（1.0=理论失效） | damage limit
              xReset 计数与损伤复位上升沿
   输出契约 : fDamageAcc 累积损伤度；iCycles 已计数全循环个数；iStackLevel 反转点栈深
              fRangeMax 已统计最大循环幅值 [µε]；xOverDamage 损伤超限锁存
              xValid 输入有效；iErrorCode 0=正常 1=非有限或参数非法 2=栈满降级
   算法说明 : 三点法判据——设栈顶三点 A,B,C，幅值 R1=|A−B|、R2=|B−C|；
              若 R2 ≥ R1 则 A→B 构成一个全循环（幅值 R1），弹出 A、B 两点；
              线性 S-N 近似取 N = fSnCoeff / R1，单循环损伤 = 1/N
   修改记录 : v1.0.0 2026-11-24 初版
   =========================================================================== *)

TYPE E_DL_FatigueDir :
(
    eDirNone := 0,   // 未定向（初始） | undirected initial
    eDirUp := 1,     // 上升段 | rising run
    eDirDown := 2    // 下降段 | falling run
);
END_TYPE

FUNCTION_BLOCK FB_DL_StrainFatigueCounter
VAR_INPUT
    fStrain : REAL;                        // 应变输入 [µε] | strain input [µε]
    fDeadBand : REAL := 5.0;               // 反转识别死区 [µε] | reversal dead band [µε]
    fSnCoeff : REAL := 500.0;              // S-N 系数（N=1 对应幅值） [µε] | sn coefficient [µε]
    fDamageLimit : REAL := 1.0;            // 损伤度限值 | damage limit
    xReset : BOOL;                         // 复位上升沿 | reset rising edge
END_VAR
VAR_OUTPUT
    fDamageAcc : REAL;                     // 累积损伤度 | accumulated damage
    iCycles : INT;                         // 已计数全循环个数 | counted full cycles
    iStackLevel : INT;                     // 反转点栈深 | reversal stack level
    fRangeMax : REAL;                      // 已统计最大循环幅值 [µε] | max counted range [µε]
    xOverDamage : BOOL;                    // 损伤超限锁存 | latched over-damage
    xValid : BOOL;                         // 输入有效标志 | inputs valid flag
    iErrorCode : INT;                      // 故障码 0=无故障 | error code
    eDirOut : E_DL_FatigueDir;             // 当前走向观测 | current direction observation
END_VAR
VAR
    _eDir : E_DL_FatigueDir := eDirNone;   // 内部走向状态 | internal direction state
    _afRev : ARRAY[1..8] OF REAL;          // 反转点栈 [µε] | reversal point stack [µε]
    _iTop : INT;                           // 栈顶下标 0=空 | stack top index
    _k : INT;                              // 前移循环下标 | shift loop index
    _fExtreme : REAL;                      // 当前走向极值 [µε] | extreme in current run [µε]
    _fPushVal : REAL;                      // 待入栈反转点 [µε] | reversal to push [µε]
    _fR1 : REAL;                           // 内层循环幅值 [µε] | inner range [µε]
    _fR2 : REAL;                           // 外层循环幅值 [µε] | outer range [µε]
    _fN : REAL;                            // 该幅值对应寿命（循环数） | life at that range
    _xPush : BOOL;                         // 本拍有待入栈反转点 | pending push flag
    _xPair : BOOL;                         // 三点配对继续标志 | pairing continue flag
    _xInit : BOOL;                         // 首拍初始化完成 | first cycle done
    _xBad : BOOL;                          // 输入非有限标志 | not-finite flag
    _xBadPar : BOOL;                       // 参数非法标志 | invalid parameter flag
    _rtReset : R_TRIG;                     // 复位上升沿 | reset rising edge
END_VAR

// ---- 无条件每周期调用：复位沿检测 ----
_rtReset(CLK := xReset);

// ---- 非有限检测 ----
_xBad := (fStrain <> fStrain) OR ((fStrain - fStrain) <> (fStrain - fStrain))
      OR (fDeadBand <> fDeadBand) OR ((fDeadBand - fDeadBand) <> (fDeadBand - fDeadBand));

// ---- 参数合法性：死区与 S-N 系数必须为正（两者都充当分母或判据） ----
_xBadPar := (fDeadBand <= 0.0) OR (fSnCoeff <= 0.0) OR (fDamageLimit <= 0.0);

// ---- 输出预置：损伤度为积分量，不做每拍清零 ----
xValid := NOT (_xBad OR _xBadPar);
iErrorCode := 0;
IF _xBad THEN
    iErrorCode := 1;
ELSIF _xBadPar THEN
    iErrorCode := 1;
END_IF

// ---- 首拍只记录极值，不产生任何循环 ----
IF NOT _xInit THEN
    _xInit := TRUE;
    _fExtreme := fStrain;
END_IF

IF xValid THEN
    // ---- 方向状态机：带死区的反转识别 ----
    _xPush := FALSE;
    _fPushVal := 0.0;
    CASE _eDir OF
        eDirNone:
            IF (fStrain - _fExtreme) > fDeadBand THEN
                _eDir := eDirUp;                       // 首次确立上升走向
                _fExtreme := fStrain;
            ELSIF (_fExtreme - fStrain) > fDeadBand THEN
                _eDir := eDirDown;                     // 首次确立下降走向
                _fExtreme := fStrain;
            END_IF

        eDirUp:
            IF fStrain > _fExtreme THEN
                _fExtreme := fStrain;                  // 刷新上升段高点
            ELSIF fStrain < (_fExtreme - fDeadBand) THEN
                _fPushVal := _fExtreme;                // 高点确认反转，待入栈
                _xPush := TRUE;
                _eDir := eDirDown;
                _fExtreme := fStrain;
            END_IF

        eDirDown:
            IF fStrain < _fExtreme THEN
                _fExtreme := fStrain;                  // 刷新下降段低点
            ELSIF fStrain > (_fExtreme + fDeadBand) THEN
                _fPushVal := _fExtreme;                // 低点确认反转，待入栈
                _xPush := TRUE;
                _eDir := eDirUp;
                _fExtreme := fStrain;
            END_IF

    ELSE
        _eDir := eDirNone;                             // 非法走向兜底重新定向
        _fExtreme := fStrain;
    END_CASE

    // ---- 入栈与三点配对 ----
    IF _xPush THEN
        IF _iTop >= 8 THEN
            // 栈满降级：丢弃最旧两点后仍继续入栈，并记录降级码
            FOR _k := 1 TO 6 DO
                _afRev[_k] := _afRev[_k + 2];
            END_FOR
            _iTop := 6;
            iErrorCode := 2;
        END_IF
        _iTop := _iTop + 1;
        _afRev[_iTop] := _fPushVal;

        _xPair := TRUE;
        WHILE _xPair AND (_iTop >= 3) DO
            _fR1 := ABS(_afRev[_iTop - 2] - _afRev[_iTop - 1]);
            _fR2 := ABS(_afRev[_iTop - 1] - _afRev[_iTop]);
            IF _fR2 >= _fR1 THEN
                // ---- 构成一个全循环，幅值 R1 ----
                IF _fR1 > 0.000001 THEN
                    _fN := fSnCoeff / _fR1;            // 分母已守卫
                    IF _fN < 1.0 THEN
                        _fN := 1.0;                    // 寿命下限 1 次，防损伤爆炸
                    END_IF
                    fDamageAcc := fDamageAcc + 1.0 / _fN;   // 分母已守卫
                    iCycles := iCycles + 1;
                    IF _fR1 > fRangeMax THEN
                        fRangeMax := _fR1;
                    END_IF
                END_IF
                // ---- 弹出 A、B 两点：剩余元素整体前移两位 ----
                FOR _k := 1 TO (_iTop - 2) DO
                    _afRev[_k] := _afRev[_k + 2];
                END_FOR
                _iTop := _iTop - 2;
            ELSE
                _xPair := FALSE;                       // 不满足判据，退出配对循环
            END_IF
        END_WHILE
    END_IF

    // ---- 损伤超限锁存与唯一解除路径 ----
    IF fDamageAcc >= fDamageLimit THEN
        xOverDamage := TRUE;
    END_IF
    IF _rtReset.Q AND NOT xOverDamage THEN
        fDamageAcc := 0.0;                             // 无锁存时复位仅清计数器
        iCycles := 0;
        iStackLevel := 0;
    ELSIF _rtReset.Q AND xOverDamage THEN
        xOverDamage := FALSE;                          // 解除路径：复位上升沿
        fDamageAcc := 0.0;
        iCycles := 0;
        fRangeMax := 0.0;
        _iTop := 0;
        _eDir := eDirNone;
        _xInit := FALSE;
    END_IF
END_IF

iStackLevel := _iTop;
eDirOut := _eDir;
END_FUNCTION_BLOCK

(* ---- FB_DL_StrainZeroDriftMon.st ---- *)
(* ===========================================================================
   组件名   : FB_DL_StrainZeroDriftMon
   分类     : DL_Device / 应变零点漂移监控
   一句话   : 空载窗口内平滑跟踪零点并累计漂移速率与总漂移量，超限锁存报警
   复杂度   : 2        版本 : v1.0.0        日期 : 2026-11-24
   开源溯源 : 无（clean-room 自研，未借鉴任何开源实现）
   输入契约 : xEnable 监控使能；fReading 当前读数 [µε]；xNoLoad 空载窗口标志
              fZeroNominal 标称零点 [µε]；fDtSec 采样周期 [s]；fWindowSec 窗口最短判定时长 [s]
              fRateLimit 漂移速率限值 [µε/min]；fAbsLimit 总漂移限值 [µε]；xReset 复位沿
   输出契约 : fZeroEst 跟踪零点 [µε]；fDriftRate 漂移速率 [µε/min]
              fDriftTotal 相对标称零点的总漂移 [µε]；fWindowSecOut 当前窗口时长 [s]
              xAlarm 超限锁存；xValid 输入有效
              iErrorCode 0=正常 1=非有限 2=参数非法 3=漂移超限
   修改记录 : v1.0.0 2026-11-24 初版
   =========================================================================== *)

FUNCTION_BLOCK FB_DL_StrainZeroDriftMon
VAR_INPUT
    xEnable : BOOL;                     // 监控使能 | monitoring enable
    fReading : REAL;                    // 当前读数 [µε] | current reading [µε]
    xNoLoad : BOOL;                     // 空载窗口标志 | no-load window flag
    fZeroNominal : REAL := 0.0;         // 标称零点 [µε] | nominal zero [µε]
    fDtSec : REAL := 0.01;              // 采样周期 [s] | sample period [s]
    fWindowSec : REAL := 30.0;          // 窗口最短判定时长 [s] | min window duration [s]
    fRateLimit : REAL := 2.0;           // 漂移速率限值 [µε/min] | drift rate limit [µε/min]
    fAbsLimit : REAL := 20.0;           // 总漂移限值 [µε] | total drift limit [µε]
    xReset : BOOL;                      // 报警复位上升沿 | alarm reset rising edge
END_VAR
VAR_OUTPUT
    fZeroEst : REAL;                    // 跟踪零点 [µε] | tracked zero [µε]
    fDriftRate : REAL;                  // 漂移速率 [µε/min] | drift rate [µε/min]
    fDriftTotal : REAL;                 // 总漂移量 [µε] | total drift [µε]
    fWindowSecOut : REAL;               // 当前窗口时长 [s] | current window duration [s]
    xAlarm : BOOL;                      // 漂移超限锁存 | latched drift alarm
    xValid : BOOL;                      // 输入有效标志 | inputs valid flag
    iErrorCode : INT;                   // 故障码 0=无故障 | error code
END_VAR
VAR
    _fDt : REAL;                        // 钳位后采样周期 [s] | clamped dt [s]
    _fWin : REAL;                       // 窗口累计时长 [s] | accumulated window [s]
    _fZeroStart : REAL;                 // 窗口起始零点 [µε] | zero at window start [µε]
    _fZero : REAL;                      // 内部跟踪零点 [µε] | internal tracked zero [µε]
    _xBad : BOOL;                       // 输入非有限标志 | not-finite flag
    _xBadPar : BOOL;                    // 参数非法标志 | invalid parameter flag
    _rtReset : R_TRIG;                  // 复位上升沿 | reset rising edge
END_VAR

// ---- 无条件每周期调用：复位沿检测 ----
_rtReset(CLK := xReset);

// ---- 非有限检测 ----
_xBad := (fReading <> fReading) OR ((fReading - fReading) <> (fReading - fReading))
      OR (fZeroNominal <> fZeroNominal) OR ((fZeroNominal - fZeroNominal) <> (fZeroNominal - fZeroNominal))
      OR (fDtSec <> fDtSec) OR ((fDtSec - fDtSec) <> (fDtSec - fDtSec));

// ---- 参数合法性 ----
_xBadPar := (fDtSec <= 0.0) OR (fWindowSec <= 0.0) OR (fRateLimit <= 0.0) OR (fAbsLimit <= 0.0);

// ---- 输出预置：报警为锁存量，不在本处清零 ----
fDriftRate := 0.0;
xValid := NOT (_xBad OR _xBadPar);
iErrorCode := 0;
IF _xBad THEN
    iErrorCode := 1;
ELSIF _xBadPar THEN
    iErrorCode := 2;
END_IF

// ---- 周期钳位 ----
_fDt := fDtSec;
IF _fDt < 0.000001 THEN
    _fDt := 0.000001;
ELSIF _fDt > 0.5 THEN
    _fDt := 0.5;
END_IF

IF xValid AND xEnable THEN
    IF xNoLoad THEN
        IF _fWin <= 0.0 THEN
            _fZeroStart := fReading;               // 窗口起点锁定零点基准
            _fZero := fReading;
        ELSE
            _fZero := _fZero + 0.05 * (fReading - _fZero);   // 指数平滑跟踪，抑制噪声
        END_IF
        _fWin := _fWin + _fDt;

        // ---- 速率计算：窗口至少满 1 s 才有意义（防除零） ----
        IF _fWin > 1.0 THEN
            fDriftRate := (_fZero - _fZeroStart) / _fWin * 60.0;   // 分母已守卫
        END_IF
    ELSE
        _fWin := 0.0;                              // 退出空载窗口即重新开始
    END_IF

    // ---- 总漂移相对标称零点 ----
    fDriftTotal := _fZero - fZeroNominal;

    // ---- 超限置位：窗口须先满最短判定时长，避免上电瞬间误报 ----
    IF (_fWin >= fWindowSec) THEN
        IF (ABS(fDriftRate) > fRateLimit) OR (ABS(fDriftTotal) > fAbsLimit) THEN
            xAlarm := TRUE;
        END_IF
    END_IF
END_IF

// ---- 报警锁存与唯一解除路径 ----
// 解除门要求 NOT xEnable，必须放在使能门控块之外评估，否则该路径永不可达
IF _rtReset.Q AND NOT xEnable THEN
    xAlarm := FALSE;
END_IF
IF xAlarm THEN
    iErrorCode := 3;
END_IF

fZeroEst := _fZero;
fWindowSecOut := _fWin;
END_FUNCTION_BLOCK

(* ---- FB_DL_TankN2BlanketCtrl.st ---- *)
//==============================================================================
// 功能块：FB_DL_TankN2BlanketCtrl ｜ 中文名称：储罐氮封压力双分程控制
// 所属子库：DL_Device ｜ 版本：v1.0.1 ｜ 兼容：CODESYS V3.5+ / TwinCAT 3 / 汇川 InoProShop
// 功能描述：储罐氮封双分程——罐压低于低压分界按比例开补氮阀位（0~100%
//           连续段），高于高压分界关量泄放；两段互斥断言（任一拍
//           NOT(fN2ChargePct > 0 AND bVentCmd)）结构性成立；分界滞环提示；
//           压力冻结/非有限判传感器断线。v1.0.1 补迟滞回差（R23 终审
//           挂账修复）：泄放段退出阈值 = fPressHiKpa - fVentHystKpa
//           （进入阈值不变，退出沿以回差带下沿为准）；补氮段审计同理
//           （进入/退出阈值分离）：退出阈值 = fPressLoKpa + fVentHystKpa，
//           两段共用同一回差带宽度语义（不新占码位）。回差非法（<= 0
//           或 >= 分界跨度）→ 故障 0357 复用并回退默认 0.2 kPa；默认仍
//           越跨度时按跨度半宽钳定（防死循环），仍报 0357。
// 开源溯源 (Origin)：道莅原创实现（参考储罐氮封系统工程惯例 分类与参数域）
// 单位表：p[kPa]（表压）/ 分界[kPa] / 阀位[%] / 延时[ms]
// 错误码表：16#0003_0184 信息级（分界点附近滞环提示，或回差带内驻留
//           提示，不置 bError）/ 16#0003_0185 预留禁用（不得挪用）/
//           16#0003_0357 故障级（分程倒置 fPressHiKpa <= fPressLoKpa、
//           回差非法 fVentHystKpa <= 0 或 >= 分界跨度，或罐压非有限
//           全关安全侧，置 bError）/ 16#0003_0358 故障级（压力冻结超窗
//           判传感器断线，置 bError）/ 16#0003_0359 故障级兜底（置
//           bError）
// 状态机：E_DL_N2BlanketState（五态：eIdle=0 / eCharging=10 / eHold=20 /
//           eVenting=30 / eFault=99），CASE 含 ELSE 兜底，ELSE 置 0359 并全关
// 边界行为：① fPressHiKpa <= fPressLoKpa → 故障 0357（分程倒置）；② 两段
//           互斥由 IF/ELSE 单源赋值结构性保证（低压段才算阀位、高压段才
//           置泄放，中间保持段两路全断）；③ 罐压非有限 → 全关（安全侧）
//           + 故障 0357 复用（R90）；④ 压力冻结超 tPressLossDelay 判断线
//           → 故障 0358；⑤ 未使能输出冻结为零并 bValid := FALSE；⑥
//           泄放退出沿 = 罐压 < fPressHiKpa - fVentHystKpa（回差带下沿），
//           补氮退出沿 = 罐压 > fPressLoKpa + fVentHystKpa（回差带上沿），
//           进入阈值两侧均不变；回差非法回退默认 0.2 kPa 仍越跨度时按
//           跨度半宽钳定并保持 0357 报警。
// 依赖收窄 (R11 留档③)：Device 不得调用 DL_Algo——分程律在本件内联实现
//           （低压段线性补氮 + 高压段开关量泄放），与 FB_DL_SplitRangeControl
//           的参数域一致性（分界点语义、0~100% 线性段）由本件头注释承担
//           验证责任，改动任一侧须复核另一侧。
// 修订历史：v1.0.0 2026-11-17 首版（R23 派单 · ROADMAP P1 §396）
//           v1.0.1 2026-11-17 R24 挂账修复：补泄放退出迟滞回差（新增
//           输入引脚 fVentHystKpa : LREAL := 0.2 [kPa]，默认非魔法数，
//           不新占码位），eVenting 退出沿以回差带下沿为准；补氮段迟滞
//           同理审计（进入/退出阈值分离，共用同一回差带宽）；回差非法
//           → 0357 复用并回退默认；0003_0184 信息级语义扩展为滞环/回差
//           驻留提示。引脚契约其余不变，枚举不变。
//==============================================================================

(*------------------------------------------------------------------------------
 * 枚举: E_DL_N2BlanketState（归属本功能块，同文件发布，全库唯一定义）
 * 含义: 氮封工作相位，每个成员在 CASE 中有且仅有一个标签。
 *-----------------------------------------------------------------------------*)
TYPE E_DL_N2BlanketState :
(
    eIdle     := 0,   // 空闲：未使能 / Idle, not enabled
    eCharging := 10,  // 补氮中：罐压低于低压分界，补氮阀位有效 / Charging, pressure below the low boundary
    eHold     := 20,  // 保持：罐压在两分界之间，两路全断 / Hold, pressure between the boundaries, both off
    eVenting  := 30,  // 泄放中：罐压达高压分界，泄放阀开 / Venting, pressure at the high boundary
    eFault    := 99   // 故障：组态非法/断线/非有限/非法状态 / Fault, illegal config, loss, non-finite or illegal state
);
END_TYPE

FUNCTION_BLOCK FB_DL_TankN2BlanketCtrl
VAR_INPUT
    fTankPressKpa   : LREAL;                // 罐压实测 [千帕]，表压 / Measured tank pressure [kPa], gauge
    fPressLoKpa     : LREAL := 0.5;         // 低压分界 [千帕]，低于此补氮 / Low boundary [kPa], charge below
    fPressHiKpa     : LREAL := 2.0;         // 高压分界 [千帕]，须 > 低压分界，达此泄放 / High boundary [kPa], must exceed the low, vent at
    fVentHystKpa    : LREAL := 0.2;         // 泄放/补氮退出迟滞回差 [千帕]，有效域 (0, 分界跨度)，v1.0.1 新增 / Vent and charge exit hysteresis [kPa], added in v1.0.1
    fN2ValveOutFb   : BOOL;                 // 补氮阀开反馈 [—] / N2 charge valve open feedback
    bEnable         : BOOL;                 // 控制使能 [—] / Control enable
    bReset          : BOOL;                 // 故障复位 [—] / Fault reset
END_VAR
VAR_OUTPUT
    fN2ChargePct    : LREAL;                // 补氮阀位 [百分数]，0~100，仅低压段有效 / N2 charge valve position [percent], 0..100, low band only
    bVentCmd        : BOOL;                 // 泄放阀指令 [—]，开关量，仅高压段 / Vent valve command, on/off, high band only
    eBlanketState   : E_DL_N2BlanketState;  // 氮封相位 [—] / Blanket phase
    eErr            : UDINT;                // 错误码，0 = 无错 / Error code, 0 = no error
    bError          : BOOL;                 // 故障级标志，仅故障级错误置位 / Fault-class flag, set only on fault-level codes
    bValid          : BOOL;                 // 输出可用标志 / Outputs usable flag
END_VAR
VAR
    fbFrozen        : TON;                  // 压力冻结判窗（断线检测），段 6 无条件刷新 [ms] / Frozen-pressure window, loss detection
    _fPressPrev     : LREAL;                // 上拍罐压快照（冻结检测基准） / Previous-scan pressure snapshot
    _bInit          : BOOL := FALSE;        // 首扫标志，初值 FALSE 取非判定 / First-scan flag, tested negated
    _bSplitBad      : BOOL;                 // 分程倒置/非有限锁存 / Inversion or non-finite latch
    _bFrozenBad     : BOOL;                 // 压力冻结锁存 / Frozen-pressure latch
    _bNearBand      : BOOL;                 // 分界滞环当拍标志 / Near-boundary flag of this scan
    _fHystEff       : LREAL;                // 生效回差带宽度 [千帕]（非法回退默认/钳定） / Effective hysteresis width [kPa]
    _bHystBad       : BOOL;                 // 回差非法锁存（0357 复用） / Illegal hysteresis latch
    _bIllegal       : BOOL;                 // 非法状态标志 / Illegal state flag
    _eState         : E_DL_N2BlanketState := E_DL_N2BlanketState.eIdle; // 当前相位 / Current phase
END_VAR
VAR CONSTANT
    DL_N2_INF       : LREAL := 1.7976931348623157E308; // LREAL 幅值上限 / LREAL magnitude ceiling
    DL_N2_LOSS_TOL  : LREAL := 1.0E-9;      // 冻结判据容差 [千帕] / Frozen detection tolerance [kPa]
    DL_N2_LOSS_WIN  : TIME  := T#5S;        // 压力冻结判窗 [ms] / Frozen-pressure window [ms]
    DL_N2_BAND_TOL  : LREAL := 0.05;        // 分界滞环提示带 [千帕] / Near-boundary notice band [kPa]
    DL_N2_HYST_DEF  : LREAL := 0.2;         // 回差带宽度默认值 [千帕]，非法时回退目标（v1.0.1） / Hysteresis default [kPa], fallback target in v1.0.1
    DL_N2_EPS       : LREAL := 1.0E-6;      // 浮点判零容差 [千帕] / Float zero tolerance [kPa]
END_VAR

(*------------------------------------------------------------------------------
 * 段 1｜每拍预置：双输出先全关（安全侧），单拍标志预清零
 *      Both outputs closed first, fail-safe, one-shot flags pre-cleared
 *-----------------------------------------------------------------------------*)
fN2ChargePct  := 0.0;                       // 补氮阀位先清（安全侧） / Charge position cleared first
bVentCmd      := FALSE;                     // 泄放指令先清（安全侧） / Vent command cleared first
eErr          := 16#0000_0000;              // 错误码每拍重算 / Error code recomputed
bError        := FALSE;                     // 故障标志每拍重算 / Fault flag recomputed
bValid        := FALSE;                     // 可用标志每拍重算 / Usable flag recomputed
_bNearBand    := FALSE;                     // 滞环标志预清零 / Near-band flag pre-cleared
_bIllegal     := FALSE;                     // 非法状态预清零 / Illegal flag pre-cleared

(*------------------------------------------------------------------------------
 * 段 2｜首扫初始化
 *      First-scan initialisation
 *-----------------------------------------------------------------------------*)
IF NOT _bInit THEN
    _eState     := E_DL_N2BlanketState.eIdle; // 相位空闲起步 / Phase starts idle
    _fPressPrev := 0.0;                     // 压力快照从零起步 / Pressure snapshot starts at zero
    _bSplitBad  := FALSE;                   // 分程锁存清零 / Inversion latch cleared
    _bFrozenBad := FALSE;                   // 冻结锁存清零 / Frozen latch cleared
    _bHystBad   := FALSE;                   // 回差锁存清零（v1.0.1） / Hysteresis latch cleared, v1.0.1
    _fHystEff   := DL_N2_HYST_DEF;          // 回差从默认起步（v1.0.1） / Hysteresis starts at the default, v1.0.1
    _bInit      := TRUE;                    // 首扫只做一次 / The first scan runs once
END_IF

(*------------------------------------------------------------------------------
 * 段 3｜组态与输入防御闸（分程倒置 / 非有限 → 0357 复用，R90）
 *      Configuration and input defense gates, code reused per R90
 *-----------------------------------------------------------------------------*)
IF (fTankPressKpa <> fTankPressKpa) OR (ABS(fTankPressKpa) > DL_N2_INF)
   OR (fPressLoKpa <> fPressLoKpa) OR (ABS(fPressLoKpa) > DL_N2_INF)
   OR (fPressHiKpa <> fPressHiKpa) OR (ABS(fPressHiKpa) > DL_N2_INF) THEN
    _bSplitBad := TRUE;                     // 非有限输入归入分程非法（安全侧全关） / Non-finite folded into the inversion fault, fail-safe closed
END_IF
IF (NOT _bSplitBad) AND (fPressHiKpa <= fPressLoKpa) THEN
    _bSplitBad := TRUE;                     // 分程倒置锁存 / Inversion latched
END_IF

(*------------------------------------------------------------------------------
 * 段 3b｜回差带宽度合法性闸（v1.0.1）：非法回退默认，默认仍越跨度按半宽钳定
 *      Hysteresis validity gate, fallback to default, half-span clamp
 *-----------------------------------------------------------------------------*)
IF (NOT _bSplitBad)
   AND ((fVentHystKpa <> fVentHystKpa) OR (ABS(fVentHystKpa) > DL_N2_INF)
        OR (fVentHystKpa <= DL_N2_LOSS_TOL)
        OR (fVentHystKpa >= (fPressHiKpa - fPressLoKpa))) THEN
    _bHystBad := TRUE;                      // 回差非法锁存（0357 复用，R90：滞环语义扩展不新占码位） / Illegal hysteresis latched
    _fHystEff := DL_N2_HYST_DEF;            // 回退默认值 / Fallback to the default
    IF _fHystEff >= (fPressHiKpa - fPressLoKpa) THEN
        _fHystEff := 0.5 * (fPressHiKpa - fPressLoKpa); // 默认仍越跨度：按跨度半宽钳定（防死循环） / Default beyond span, clamped to half span
    END_IF
ELSIF NOT _bSplitBad THEN
    _fHystEff := fVentHystKpa;              // 合法回差原值生效 / Legal hysteresis applied as-is
ELSE
    _fHystEff := DL_N2_HYST_DEF;            // 分程已非法：回差取默认（不重复报码，R90） / Split already illegal, default width, no duplicate code
END_IF

(*------------------------------------------------------------------------------
 * 段 4｜压力冻结检测：罐压与上拍差 < 容差持续超窗 → 判传感器断线
 *      Frozen-pressure detection, loss suspected beyond the window
 *-----------------------------------------------------------------------------*)
fbFrozen(IN := bEnable AND (NOT _bSplitBad)
             AND (ABS(fTankPressKpa - _fPressPrev) < DL_N2_LOSS_TOL), PT := DL_N2_LOSS_WIN); // 压力冻结判窗 / Frozen-pressure window
_fPressPrev := fTankPressKpa;               // 快照推进 / Snapshot advanced
IF fbFrozen.Q THEN
    _bFrozenBad := TRUE;                    // 断线锁存（安全侧全关） / Loss latched, fail-safe closed
END_IF
IF bReset THEN
    _bFrozenBad := FALSE;                   // 复位清冻结锁存 / Reset clears the frozen latch
    _bHystBad   := FALSE;                   // 复位清回差非法锁存（v1.0.1） / Reset clears the hysteresis latch, v1.0.1
END_IF

(*------------------------------------------------------------------------------
 * 段 5｜相位机与分程律内联（互斥断言：低压段才算阀位、高压段才置泄放）
 *      Phase machine and the inline split-range law, mutually exclusive
 *-----------------------------------------------------------------------------*)
IF (NOT bEnable) OR _bSplitBad OR _bFrozenBad THEN
    _eState := E_DL_N2BlanketState.eFault;  // 未使能或异常转故障态（全关） / Not enabled or anomaly, fault with all closed
ELSE
CASE _eState OF

    E_DL_N2BlanketState.eIdle:             // 空闲：使能即进保持
        IF bEnable THEN
            _eState := E_DL_N2BlanketState.eHold; // 进保持 / To hold
        END_IF

    E_DL_N2BlanketState.eHold:             // 保持：分界判定进补氮或泄放
        IF fTankPressKpa <= fPressLoKpa THEN
            _eState := E_DL_N2BlanketState.eCharging; // 进补氮 / To charging
        ELSIF fTankPressKpa >= fPressHiKpa THEN
            _eState := E_DL_N2BlanketState.eVenting; // 进泄放 / To venting
        END_IF
        IF (ABS(fTankPressKpa - fPressLoKpa) < DL_N2_BAND_TOL)
           OR (ABS(fTankPressKpa - fPressHiKpa) < DL_N2_BAND_TOL) THEN
            _bNearBand := TRUE;             // 分界滞环提示 / Near-boundary notice
        END_IF

    E_DL_N2BlanketState.eCharging:         // 补氮：罐压超回差带上沿（v1.0.1 阈值分离）即回保持
        IF fTankPressKpa > (fPressLoKpa + _fHystEff) THEN
            _eState := E_DL_N2BlanketState.eHold; // 回保持 / Back to hold
        END_IF

    E_DL_N2BlanketState.eVenting:          // 泄放：罐压跌破回差带下沿（v1.0.1 退出沿）即回保持
        IF fTankPressKpa < (fPressHiKpa - _fHystEff) THEN
            _eState := E_DL_N2BlanketState.eHold; // 回保持 / Back to hold
        END_IF

    E_DL_N2BlanketState.eFault:            // 故障：复位沿且原因消失回保持
        IF bReset AND (NOT _bSplitBad) AND (NOT _bFrozenBad) AND bEnable THEN
            _eState := E_DL_N2BlanketState.eHold; // 回保持 / Back to hold
        END_IF

    ELSE                                   // 非法状态兜底（R21：CASE 必带 ELSE）
        _bIllegal := TRUE;                 // 标记非法状态 / Flag the illegal state
        _eState   := E_DL_N2BlanketState.eFault; // 回故障态（全关） / Back to fault, all closed
END_CASE
END_IF

(*------------------------------------------------------------------------------
 * 段 6｜输出置位：IF/ELSE 单源赋值，两段互斥结构性成立
 *      Output assignment, mutual exclusion holds structurally
 *-----------------------------------------------------------------------------*)
CASE _eState OF
    E_DL_N2BlanketState.eCharging:         // 补氮段：阀位按低压段深度线性（0~100%） / Charging: position linear in the low band
        IF ABS(fPressLoKpa) > DL_N2_EPS THEN
            fN2ChargePct := MIN(MAX((fPressLoKpa - fTankPressKpa) / fPressLoKpa, 0.0), 1.0) * 100.0; // 补氮阀位 [百分数]，分母已闸 / Charge position, denominator gated
        ELSE
            fN2ChargePct := 100.0;          // 低压分界为 0：全开补氮（退化域防御） / Zero boundary, full charge
        END_IF
        bVentCmd := FALSE;                  // 泄放指令断（互斥断言） / Vent command off, mutually exclusive
    E_DL_N2BlanketState.eVenting:          // 泄放段：泄放开、补氮全关 / Venting: vent on, charge fully closed
        fN2ChargePct := 0.0;               // 补氮全关 / Charge fully closed
        bVentCmd := TRUE;                  // 泄放指令开 / Vent command on
    ELSE                                   // 其余相两路全关（含保持/故障） / Otherwise both closed, hold and fault
        fN2ChargePct := 0.0;               // 补氮全关 / Charge fully closed
        bVentCmd := FALSE;                 // 泄放指令断 / Vent command off
END_CASE
eBlanketState := _eState;                   // 相位出口 / Phase outlet

(*------------------------------------------------------------------------------
 * 段 7｜码位出口
 *      Code outlet
 *-----------------------------------------------------------------------------*)
IF _bIllegal THEN
    eErr   := 16#0003_0359;                 // 故障级：状态机兜底 / Fault: fallback
    bError := TRUE;                         // 置故障标志 / Raise the fault flag
ELSIF _bSplitBad OR _bFrozenBad OR _bHystBad THEN
    IF _bFrozenBad AND (NOT _bSplitBad) AND (NOT _bHystBad) THEN
        eErr   := 16#0003_0358;             // 故障级：压力冻结判断线 / Fault: frozen pressure, loss suspected
    ELSE
        eErr   := 16#0003_0357;             // 故障级：分程倒置/回差非法/非有限（R90 复用） / Fault: inversion, illegal hysteresis or non-finite, code reused
    END_IF
    bError := TRUE;                         // 置故障标志 / Raise the fault flag
ELSIF _bNearBand THEN
    eErr := 16#0003_0184;                   // 信息级：分界滞环提示 / Info: near-boundary notice
END_IF

bValid := (NOT bError) AND bEnable AND (_eState <> E_DL_N2BlanketState.eIdle); // 空闲/故障/未使能输出不可用 / Outputs unusable in idle, fault or disabled
END_FUNCTION_BLOCK

(* ---- FB_DL_TcChannelScanDiag.st ---- *)
(*==============================================================================
 * 组件名称 (Component)  : FB_DL_TcChannelScanDiag
 * 所属子库 (Sublibrary) : DL_Device
 * 当前版本 (Version)    : 1.0.0
 * 兼容性   (Platform)   : CODESYS 3.5+ / TwinCAT 3 / 汇川 InoProShop / 施耐德 Machine Expert
 *                         仅依赖 Standard.library（R_TRIG / ABS），零厂商私有库
 * 功能描述 (Function)   : 多路热电偶断偶/反接/漂移诊断，逐通道轮询扫描（每拍扫一路，8 路一轮 8 拍）。
 *                         三类特征按优先级判定（优先级即归因优先级，先断偶后反接再漂移）：
 *                           ① 断偶 = 超量程特征：读数高于量程上限或低于量程下限（开路时前端
 *                              常表现为满量程上冲或极度负偏，故用双侧超量程判，不只判高侧）；
 *                           ② 反接 = 负向特征：读数低于 fNegThresh（明显负温，正常工况不会出现）；
 *                           ③ 漂移 = 慢变趋势特征：读数与慢变基线（EMA，系数 fDriftAlpha）之差
 *                              持续超 fDriftBand。用"基线 vs 瞬时"而非"两拍差分"，因为两拍差分
 *                              会被噪声主导；EMA 基线滤掉噪声只留趋势，正是慢变趋势的定义。
 *                         故障码按通道编码：每通道一个 ENUM 槽（aeFault[i]），另有 nFaultMask
 *                         位掩码（bit i = 通道 i 有故障）供 HMI 一字节查看。**不占用全局事件码段**。
 *                         故障为逐通道锁存，清除路径：bReset 上升沿（全清）——单通道清不在本件
 *                         （单通道清应由上层在换传感器后整体复位，避免"故障码还在但传感器已换"
 *                         的台账错乱）。
 * 接口     (Interface)  : 输入 afTempC 8 路温度（VAR_IN_OUT，本件只读）、nChannelCount 实际通道数
 *                         （2..8）、fRangeMin / fRangeMax 量程、fNegThresh 反接负向阈（工程单位）、
 *                         fDriftBand 漂移带、fDriftAlpha 基线 EMA 系数（0..1）、bReset 复位；
 *                         输出 aeFault 逐通道故障、nFaultMask 通道位掩码、bAnyFault 任一通道故障、
 *                         nScanIdx 当前扫描通道号、fLastValue 当拍扫描通道读数、eState / bError。
 * 边界     (Boundary)   : ① **属主边界（写死）：本件只诊断传感器链路（断偶/反接/漂移），
 *                         不做温度补偿、不参与温控回路、不判超温**。超温保护属温控/安全链；
 *                         把断偶诊断塞进超温保护会让"传感器坏了"与"真超温"混为一谈。
 *                         ② 组态闸：nChannelCount < 2 或 > 8（越 ARRAY 边界，缺此即数组越界读）、
 *                         fRangeMin >= fRangeMax（量程倒置）、fNegThresh >= fRangeMin
 *                         （反接阈落在量程内会把正常低温误判反接）、fDriftBand <= 0.0、
 *                         fDriftAlpha <= 0.0 或 >= 1.0（EMA 系数必须开区间）、任一输入 NaN
 *                         → 故障锁存，全部通道停止判定（不宣称），bError 置位。
 *                         ③ 轮询用 _nIdx 自增取模，绝不越界（先钳再取模双保险）。
 *                         ④ 单枚 R_TRIG（bReset）段 0 无条件周期刷新；无 TON，故无跨相复位问题。
 *                         ⑤ 故障相迁出唯一路径 = bReset 上升沿（R228B）。
 *                         ⑥ 零全局耦合（无 GVL / 无 VAR_EXTERNAL / 无物理地址）。
 * 分工声明 (Scope)      : 与 `FB_DL_AnalogScaleEx`（模拟量标定换算）分工——那件把原始码值换成
 *                         工程单位，本件在工程单位域做**链路健康诊断**。二者串接顺序固定：
 *                         先换算后诊断（断偶判据依赖量程，量程是工程单位概念）。
 * 来源标签 (Source Tag) : T2-6 ◐（开源参考：热电偶断线/反接诊断特征参数域，零代码行复制）
 * 解除式   (Release)    : bReset 上升沿 ∧ 组态合法 → 全通道故障表清零、基线表清零（重新起 EMA）。
 *                         自证可满足：复位为外部动作，不受逐通道锁存门控。
 * 码表     (Codes)      : 本件**不占用任何全局数字码位**。故障以"逐通道 ENUM + 通道位掩码"
 *                         表达（ENUM 成员是通道内的故障种类，不是全局事件码）；数字码位待
 *                         主控收口阶段统一派号。
 * 红线自检 (Redline)    : R1 ✓ 零 GVL/VAR_EXTERNAL ｜ R2 ✓ 零 %I/%Q/%M ｜ R3 ✓ 纯 IEC 61131-3
 *                         R4 ✓ 数组边界闸 + EMA 开区间闸 + 量程几何闸 + NaN 闸
 *                         R5 ✓ 声明逐行同行双语注释 ｜ R6 ✓ ENUM+CASE 含 ELSE
 *                         R7 ✓ R_TRIG 段 0 无条件刷新
 * 修订历史 (Revision)   : 2026-11-19  v1.0.0  R46 首版（批次 3 · 序号 13）
 *==============================================================================*)

TYPE E_DL_TcdFault :
(
    eOk      := 0,    // 通道健康 / Channel healthy
    eOpen    := 10,   // 断偶（超量程特征） / Open thermocouple, out-of-range signature
    eReverse := 20,   // 反接（负向特征） / Reversed polarity, negative signature
    eDrift   := 30,   // 漂移（慢变趋势特征） / Drift, slow-trend signature
    eCfg     := 90    // 组态/输入非法，通道未判定 / Configuration or input illegal, channel not judged
);
END_TYPE

TYPE E_DL_TcdState :
(
    eIdle  := 0,    // 首轮扫描未完成 / First scan round not complete
    eRun   := 10,   // 轮询诊断运行相 / Round-robin diagnosis running
    eFault := 90    // 组态故障相 / Configuration fault phase
);
END_TYPE

FUNCTION_BLOCK FB_DL_TcChannelScanDiag
VAR_IN_OUT
    afTempC : ARRAY[0..7] OF REAL;      // 8 路温度（本件只读，按 nChannelCount 截取） [°C] / Eight channels, read-only here [degC]
END_VAR
VAR_INPUT
    nChannelCount : INT := 8;           // 实际通道数，域 2..8 / Active channel count, 2..8
    fRangeMin     : REAL := -50.0;      // 量程下限，域 < fRangeMax [°C] / Range lower bound, < upper [degC]
    fRangeMax     : REAL := 400.0;      // 量程上限，域 > fRangeMin [°C] / Range upper bound, > lower [degC]
    fNegThresh    : REAL := -20.0;      // 反接负向阈，域 < fRangeMin [°C] / Reverse-polarity threshold, < range lower [degC]
    fDriftBand    : REAL := 5.0;        // 漂移带（读数与基线之差），域 > 0.0 [°C] / Drift band, > 0.0 [degC]
    fDriftAlpha   : REAL := 0.01;       // 基线 EMA 系数，域 (0, 1) 开区间 [-] / Baseline EMA coefficient, open interval (0,1)
    bReset        : BOOL := FALSE;      // 复位，上升沿清全部通道故障 [-] / Reset, rising edge clears all channel faults
END_VAR
VAR_OUTPUT
    aeFault    : ARRAY[0..7] OF E_DL_TcdFault;   // 逐通道故障出口 [-] / Per-channel fault outlet
    nFaultMask : BYTE;                  // 通道位掩码：bit i = 通道 i 有故障 [-] / Channel bit mask, bit i = channel i faulty
    bAnyFault  : BOOL;                  // 任一通道故障（锁存） [-] / Any channel faulty, latched
    nScanIdx   : INT;                   // 本拍扫描的通道号 [通道] / Channel scanned this scan
    fLastValue : REAL;                  // 本拍扫描通道的读数 [°C] / Reading of the scanned channel [degC]
    eState     : E_DL_TcdState;         // 状态出口 [-] / State outlet
    bError     : BOOL;                  // 故障标志（任一通道故障或组态非法） [-] / Error flag
END_VAR
VAR
    _eState   : E_DL_TcdState := E_DL_TcdState.eIdle;    // 内部相位（CASE 唯一写入目标） / Internal phase
    rtReset   : R_TRIG;                 // 复位沿实例，段 0 无条件调用 / Reset edge instance
    _afBase   : ARRAY[0..7] OF REAL;    // 逐通道慢变基线（EMA，锁存量） [°C] / Per-channel slow baseline, latched [degC]
    _abInit   : ARRAY[0..7] OF BOOL;    // 逐通道基线已初始化标记（锁存量） / Per-channel baseline initialised flag
    _aeFault  : ARRAY[0..7] OF E_DL_TcdFault;   // 逐通道故障锁存表（锁存量） / Per-channel latched fault table
    _nIdx     : INT;                    // 轮询索引（锁存量） / Round-robin index, latched
    _nRound   : UDINT;                  // 已完成扫描次数（锁存量） / Completed scan rounds, latched
    _bAny     : BOOL;                   // 任一通道故障锁存位（锁存量） / Latched any-fault bit
    _bCfgBad  : BOOL;                   // 组态非法当拍量 [-] / Illegal configuration this scan
    _bNonFin  : BOOL;                   // 阈值非法当拍量 [-] / Illegal threshold this scan
    _fVal     : REAL;                   // 本拍扫描通道读数（已过边界钳位的索引取值） [°C] / Scanned channel value, index guaranteed in range
    _fDev     : REAL;                   // 读数与基线之差 [°C] / Deviation from the baseline [°C]
    _i        : INT;                    // 掩码重建索引 / Mask rebuild index
    _nSh      : INT;                    // 移位量归一后副本（0..7，禁 SHL 越位宽） [位] / Normalised shift amount, 0..7
END_VAR
VAR CONSTANT
    DL_TCD_MAXN  : INT := 8;        // 通道容量（与 ARRAY 上界一致） [通道] / Channel capacity matching the array bounds
    DL_TCD_MINN  : INT := 2;        // 最少通道数 [通道] / Minimum channel count
    DL_TCD_BIT   : BYTE := 16#01;   // 掩码左移基元 [位] / Mask shift primitive
END_VAR

(* —— 段 0：判据派生 + 复位沿无条件周期刷新 —— *)
_bNonFin := (fRangeMin <> fRangeMin) OR (fRangeMax <> fRangeMax)         // NaN 自反判（判等禁令唯一例外） / NaN self-reflexive tests
         OR (fNegThresh <> fNegThresh) OR (fDriftBand <> fDriftBand)
         OR (fDriftAlpha <> fDriftAlpha);
_bCfgBad := (nChannelCount < DL_TCD_MINN) OR (nChannelCount > DL_TCD_MAXN)   // 通道数越 ARRAY 边界闸 / Channel count against array bounds
         OR (fRangeMin >= fRangeMax)                                         // 量程倒置闸 / Range inversion gate
         OR (fNegThresh >= fRangeMin)                                        // 反接阈必须低于量程下限（否则误判低温） / Reverse threshold must lie below the range
         OR (fDriftBand <= 0.0)                                              // 漂移带须为正 / Drift band must be positive
         OR (fDriftAlpha <= 0.0) OR (fDriftAlpha >= 1.0)                     // EMA 系数开区间闸 / EMA coefficient open-interval gate
         OR _bNonFin;                                                        // 非有限 / Non-finite
rtReset(CLK := bReset);                                                     // 复位沿，每拍必调（R228A） / Reset edge, every scan

(* —— 段 1：单拍量预清零（锁存量 _aeFault/_afBase/_abInit/_nIdx/_nRound/_bAny 不入清单，R107） —— *)
bAnyFault  := FALSE;        // 任一故障出口预清 / Any-fault preset
nScanIdx   := 0;            // 扫描索引出口预清 / Scan index preset
fLastValue := 0.0;          // 读数出口预清 / Value preset
bError     := FALSE;        // 故障标志预清（R45 配对） / Error flag preset

(* —— 段 2：复位沿 + 组态闸 —— *)
IF rtReset.Q THEN
    FOR _i := 0 TO DL_TCD_MAXN - 1 DO
        _aeFault[_i] := E_DL_TcdFault.eOk;      // 全通道故障清 / Clear every channel fault
        _abInit[_i]  := FALSE;                  // 基线标记清（重新起 EMA） / Baseline flags cleared, EMA restarts
        _afBase[_i]  := 0.0;                    // 基线清 / Baselines cleared
    END_FOR
    _bAny   := FALSE;                           // 任一故障锁存清 / Clear the any-fault latch
    _nIdx   := 0;                               // 轮询索引归零 / Round-robin index cleared
    _nRound := 0;                               // 扫描轮次归零 / Round counter cleared
    IF _eState = E_DL_TcdState.eFault THEN
        _eState := E_DL_TcdState.eIdle;         // 故障相迁出（R228B） / Leave fault phase
    END_IF
END_IF
IF _bCfgBad THEN
    _eState := E_DL_TcdState.eFault;            // 组态非法入故障相 / Enter fault phase
    FOR _i := 0 TO DL_TCD_MAXN - 1 DO
        _aeFault[_i] := E_DL_TcdFault.eCfg;     // 全通道标"未判定"（不得伪报健康） / Mark every channel as not judged
    END_FOR
END_IF

(* —— 段 3：轮询索引钳位（先钳后取模，双保险防越界） —— *)
IF _nIdx < 0 THEN
    _nIdx := 0;                                 // 负索引钳位 / Clamp a negative index
END_IF
IF _nIdx > DL_TCD_MAXN - 1 THEN
    _nIdx := 0;                                 // 超上界回卷 / Wrap above the upper bound
END_IF
IF (NOT _bCfgBad) AND (_nIdx >= nChannelCount) THEN
    _nIdx := 0;                                 // 越过实际通道数回卷 / Wrap at the active channel count
END_IF

(* —— 段 4：单通道扫描判定（本拍只判一路，8 路一轮） —— *)
IF NOT _bCfgBad THEN
    _fVal := afTempC[_nIdx];                    // 索引已在段 3 钳位，取值为安全读 / Index already clamped
    nScanIdx   := _nIdx;                        // 扫描通道出口 / Scanned channel outlet
    fLastValue := _fVal;                        // 读数出口 / Value outlet
    IF (_fVal <> _fVal) THEN
        _aeFault[_nIdx] := E_DL_TcdFault.eCfg;  // 读数 NaN：该路标未判定（最可能是通道配置错） / NaN reading marks the channel not judged
    ELSIF (_fVal > fRangeMax) OR (_fVal < fRangeMin) THEN
        _aeFault[_nIdx] := E_DL_TcdFault.eOpen; // 超量程 = 断偶特征（双侧判） / Out of range on either side means open
    ELSIF _fVal < fNegThresh THEN
        _aeFault[_nIdx] := E_DL_TcdFault.eReverse;  // 负向超反接阈 = 反接特征 / Beyond the negative threshold means reversed
    ELSE
        IF _abInit[_nIdx] = FALSE THEN
            _afBase[_nIdx] := _fVal;            // 基线初始化（首读直接落盘） / Initialise the baseline with the first reading
            _abInit[_nIdx] := TRUE;             // 标记已初始化 / Mark initialised
        ELSE
            _fDev := _fVal - _afBase[_nIdx];    // 读数与基线之差 / Deviation from the baseline
            IF ABS(_fDev) > fDriftBand THEN
                _aeFault[_nIdx] := E_DL_TcdFault.eDrift;    // 慢变趋势超带 = 漂移特征 / Slow deviation beyond the band means drift
            ELSIF _aeFault[_nIdx] = E_DL_TcdFault.eDrift THEN
                _aeFault[_nIdx] := E_DL_TcdFault.eOk;       // 回到带内即清该路漂移（漂移是缓变，允许自愈） / Back inside clears drift on this channel
            END_IF
            _afBase[_nIdx] := _afBase[_nIdx] + (fDriftAlpha * _fDev);   // EMA 基线跟随（系数已闸） / EMA baseline update
        END_IF
    END_IF
    _nIdx := _nIdx + 1;                         // 索引前进 / Advance the index
    IF _nIdx >= nChannelCount THEN
        _nIdx := 0;                             // 到通道数回卷 / Wrap at the active count
        _nRound := _nRound + 1;                 // 一轮完成 / One round completed
    END_IF
END_IF

(* —— 段 5：掩码与汇总（由逐通道表重建，不独立维护，杜绝两处不一致） —— *)
nFaultMask := 16#00;                            // 掩码每拍重建 / Mask rebuilt each scan
FOR _i := 0 TO DL_TCD_MAXN - 1 DO
    IF (_i < nChannelCount) AND (_aeFault[_i] <> E_DL_TcdFault.eOk) THEN
        _nSh := _i;                                           // 移位量归一：先落副本再钳 / Normalise the shift amount first
        IF _nSh < 0 THEN
            _nSh := 0;                                        // 下界钳 / Lower clamp
        END_IF
        IF _nSh > 7 THEN
            _nSh := 7;                                        // 上界钳（BYTE 位宽 8，禁 SHL 越位宽） / Upper clamp, never shift past the BYTE width
        END_IF
        nFaultMask := nFaultMask OR SHL(DL_TCD_BIT, INT_TO_BYTE(_nSh));   // 位 i 置（移位量已归一到 0..7） / Set bit i with the shift amount normalised
        _bAny := TRUE;                                        // 任一故障锁存 / Latch the any-fault bit
    END_IF
END_FOR

(* —— 段 6：锁存相位迁移闸 —— *)
IF _bCfgBad THEN
    _bAny := TRUE;                              // 组态非法也算"有故障"（对外不宣称健康） / Illegal config counts as faulty
END_IF
IF _bAny AND (_eState <> E_DL_TcdState.eFault) AND _bCfgBad THEN
    _eState := E_DL_TcdState.eFault;            // 组态型故障入故障相 / Configuration fault enters the fault phase
END_IF

(* —— 段 7：相位机（ENUM 全成员显式标签 + ELSE 兜底，R128） —— *)
CASE _eState OF

E_DL_TcdState.eIdle:
    IF _bCfgBad THEN                            // 出口 1：组态非法 / Illegal configuration
        _eState := E_DL_TcdState.eFault;
    ELSIF _nRound >= 1 THEN                     // 出口 2：完成至少一轮，全通道已有结论 / At least one round done
        _eState := E_DL_TcdState.eRun;
    END_IF

E_DL_TcdState.eRun:
    IF _bCfgBad THEN                            // 出口 1：组态转非法 / Configuration went illegal
        _eState := E_DL_TcdState.eFault;
    ELSIF rtReset.Q THEN                        // 出口 2：复位回等待相 / Reset back to idle
        _eState := E_DL_TcdState.eIdle;
    END_IF

E_DL_TcdState.eFault:
    IF rtReset.Q AND (NOT _bCfgBad) THEN        // 出口：复位且组态已合法才迁出（R228B） / Reset with legal config
        _eState := E_DL_TcdState.eIdle;
    END_IF

ELSE
    _eState := E_DL_TcdState.eFault;            // 非法相位兜底 / Illegal-phase fallback
    bError  := TRUE;                            // 故障标志 / Error flag

END_CASE

(* —— 段 8：出口单点映射（逐通道表整体回放 + 汇总位同源，R191） —— *)
FOR _i := 0 TO DL_TCD_MAXN - 1 DO
    aeFault[_i] := _aeFault[_i];                // 逐通道故障回放 / Per-channel fault replay
END_FOR
bAnyFault := _bAny;                             // 任一故障与锁存同源 / Any-fault from latch
bError    := _bAny OR (_eState = E_DL_TcdState.eFault);    // 故障标志 = 任一故障或组态故障 / Error = any fault or config fault
eState    := _eState;                           // 状态出口 / State outlet

END_FUNCTION_BLOCK
